(* IEC 61131-3 sources: plc-st-coding-agent/progress/evidence/f14_v6_public_pilot_20261112/jobs/custom_deepseek-v4pro, 34 files *)

(* ---- public-easy-01.candidate_01.st ---- *)
(* ENGINEERING_CONTRACT
States: 0 Idle, 1 Cleaning, 2 Filling, 3 Capping, 4 Packing, 5 Complete.
Activation: bottleSensor rising edge in Idle -> Cleaning. Cleaning holds Pump_Motor until cleaningConfirmButton rising edge.
cleaningConfirmButton in Cleaning -> Filling. fillingConfirmButton in Filling -> Capping.
cappingConfirmButton in Capping -> Packing. packingConfirmButton in Packing -> Complete.
finishedButton in Complete -> Idle and resets all outputs.
Outputs active only in matching state: Pump_Motor/Cleaning, Filling_Valve/Filling,
Capping_Machine/Capping, Packing_Machine/Packing, Completion_Light/Complete.
Unspecified: simultaneous inputs in one scan resolve by current state only.
*)

(* CONTRACT_RULES [] *)

FUNCTION_BLOCK AutomatedFillingLine
VAR_INPUT
    bottleSensor : BOOL;
    cleaningConfirmButton : BOOL;
    fillingConfirmButton : BOOL;
    cappingConfirmButton : BOOL;
    packingConfirmButton : BOOL;
    finishedButton : BOOL;
END_VAR
VAR_OUTPUT
    Pump_Motor : BOOL;
    Filling_Valve : BOOL;
    Capping_Machine : BOOL;
    Packing_Machine : BOOL;
    Completion_Light : BOOL;
END_VAR
VAR
    state : INT := 0;
    tmp_nextState : INT := 0;

    tmp_lastBottle : BOOL := FALSE;
    tmp_lastCleaning : BOOL := FALSE;
    tmp_lastFilling : BOOL := FALSE;
    tmp_lastCapping : BOOL := FALSE;
    tmp_lastPacking : BOOL := FALSE;
    tmp_lastFinished : BOOL := FALSE;

    tmp_bottleRise : BOOL;
    tmp_cleaningRise : BOOL;
    tmp_fillingRise : BOOL;
    tmp_cappingRise : BOOL;
    tmp_packingRise : BOOL;
    tmp_finishedRise : BOOL;
END_VAR

(* Rising edge detection *)
tmp_bottleRise := bottleSensor AND NOT tmp_lastBottle;
tmp_lastBottle := bottleSensor;

tmp_cleaningRise := cleaningConfirmButton AND NOT tmp_lastCleaning;
tmp_lastCleaning := cleaningConfirmButton;

tmp_fillingRise := fillingConfirmButton AND NOT tmp_lastFilling;
tmp_lastFilling := fillingConfirmButton;

tmp_cappingRise := cappingConfirmButton AND NOT tmp_lastCapping;
tmp_lastCapping := cappingConfirmButton;

tmp_packingRise := packingConfirmButton AND NOT tmp_lastPacking;
tmp_lastPacking := packingConfirmButton;

tmp_finishedRise := finishedButton AND NOT tmp_lastFinished;
tmp_lastFinished := finishedButton;

(* Compute next state from current state and relevant rising edges *)
tmp_nextState := state;
CASE state OF
    0: (* Idle *)
        IF tmp_bottleRise THEN
            tmp_nextState := 1;
        END_IF;
    1: (* Cleaning *)
        IF tmp_cleaningRise THEN
            tmp_nextState := 2;
        END_IF;
    2: (* Filling *)
        IF tmp_fillingRise THEN
            tmp_nextState := 3;
        END_IF;
    3: (* Capping *)
        IF tmp_cappingRise THEN
            tmp_nextState := 4;
        END_IF;
    4: (* Packing *)
        IF tmp_packingRise THEN
            tmp_nextState := 5;
        END_IF;
    5: (* Complete *)
        IF tmp_finishedRise THEN
            tmp_nextState := 0;
        END_IF;
    ELSE
        tmp_nextState := 0;
END_CASE;
state := tmp_nextState;

(* Output assignment for current state *)
Pump_Motor := FALSE;
Filling_Valve := FALSE;
Capping_Machine := FALSE;
Packing_Machine := FALSE;
Completion_Light := FALSE;

CASE state OF
    1:
        Pump_Motor := TRUE;
    2:
        Filling_Valve := TRUE;
    3:
        Capping_Machine := TRUE;
    4:
        Packing_Machine := TRUE;
    5:
        Completion_Light := TRUE;
END_CASE;

END_FUNCTION_BLOCK

(* ---- public-easy-01.candidate_02.st ---- *)
(* ENGINEERING_CONTRACT
States: 0 Idle, 1 Cleaning, 2 Filling, 3 Capping, 4 Packing, 5 Complete.
Activation: bottleSensor rising edge in Idle -> Cleaning. Pump_Motor is latched ON by bottleSensor rising edge and latched OFF by finishedButton rising edge (per PUB003 "continues to work" interpreted as retention until process reset).
cleaningConfirmButton rising edge in Cleaning -> Filling. fillingConfirmButton rising edge in Filling -> Capping.
cappingConfirmButton rising edge in Capping -> Packing. packingConfirmButton rising edge in Packing -> Complete.
finishedButton rising edge in Complete -> Idle and resets all outputs (including Pump_Motor).
Outputs active only in matching state: Filling_Valve/Filling, Capping_Machine/Capping, Packing_Machine/Packing, Completion_Light/Complete.
Pump_Motor is NOT state-dependent; it remains true from bottle detection until finishedButton resets.
Unspecified: simultaneous inputs in one scan resolve by current state only; finishedButton outside Complete resets Pump_Motor as a global reset.
*)

(* CONTRACT_RULES [
  {"kind": "hold_until_reset", "output": "Pump_Motor", "set_input": "bottleSensor", "reset_input": "finishedButton"}
] *)

FUNCTION_BLOCK AutomatedFillingLine
VAR_INPUT
    bottleSensor : BOOL;
    cleaningConfirmButton : BOOL;
    fillingConfirmButton : BOOL;
    cappingConfirmButton : BOOL;
    packingConfirmButton : BOOL;
    finishedButton : BOOL;
END_VAR
VAR_OUTPUT
    Pump_Motor : BOOL;
    Filling_Valve : BOOL;
    Capping_Machine : BOOL;
    Packing_Machine : BOOL;
    Completion_Light : BOOL;
END_VAR
VAR
    state : INT := 0;
    pumpLatch : BOOL := FALSE;

    tmp_nextState : INT := 0;

    tmp_lastBottle : BOOL := FALSE;
    tmp_lastCleaning : BOOL := FALSE;
    tmp_lastFilling : BOOL := FALSE;
    tmp_lastCapping : BOOL := FALSE;
    tmp_lastPacking : BOOL := FALSE;
    tmp_lastFinished : BOOL := FALSE;

    tmp_bottleRise : BOOL;
    tmp_cleaningRise : BOOL;
    tmp_fillingRise : BOOL;
    tmp_cappingRise : BOOL;
    tmp_packingRise : BOOL;
    tmp_finishedRise : BOOL;
END_VAR

(* Rising edge detection *)
tmp_bottleRise := bottleSensor AND NOT tmp_lastBottle;
tmp_lastBottle := bottleSensor;

tmp_cleaningRise := cleaningConfirmButton AND NOT tmp_lastCleaning;
tmp_lastCleaning := cleaningConfirmButton;

tmp_fillingRise := fillingConfirmButton AND NOT tmp_lastFilling;
tmp_lastFilling := fillingConfirmButton;

tmp_cappingRise := cappingConfirmButton AND NOT tmp_lastCapping;
tmp_lastCapping := cappingConfirmButton;

tmp_packingRise := packingConfirmButton AND NOT tmp_lastPacking;
tmp_lastPacking := packingConfirmButton;

tmp_finishedRise := finishedButton AND NOT tmp_lastFinished;
tmp_lastFinished := finishedButton;

(* Pump latch: set on bottle detection, reset on finished button *)
IF tmp_bottleRise THEN
    pumpLatch := TRUE;
END_IF;
IF tmp_finishedRise THEN
    pumpLatch := FALSE;
END_IF;
Pump_Motor := pumpLatch;

(* Compute next state from current state and relevant rising edges *)
tmp_nextState := state;
CASE state OF
    0: (* Idle *)
        IF tmp_bottleRise THEN
            tmp_nextState := 1;
        END_IF;
    1: (* Cleaning *)
        IF tmp_cleaningRise THEN
            tmp_nextState := 2;
        END_IF;
    2: (* Filling *)
        IF tmp_fillingRise THEN
            tmp_nextState := 3;
        END_IF;
    3: (* Capping *)
        IF tmp_cappingRise THEN
            tmp_nextState := 4;
        END_IF;
    4: (* Packing *)
        IF tmp_packingRise THEN
            tmp_nextState := 5;
        END_IF;
    5: (* Complete *)
        IF tmp_finishedRise THEN
            tmp_nextState := 0;
        END_IF;
    ELSE
        tmp_nextState := 0;
END_CASE;
state := tmp_nextState;

(* Output assignment for state-dependent outputs (excluding Pump_Motor) *)
Filling_Valve := FALSE;
Capping_Machine := FALSE;
Packing_Machine := FALSE;
Completion_Light := FALSE;

CASE state OF
    2:
        Filling_Valve := TRUE;
    3:
        Capping_Machine := TRUE;
    4:
        Packing_Machine := TRUE;
    5:
        Completion_Light := TRUE;
END_CASE;

END_FUNCTION_BLOCK

(* ---- public-easy-01.candidate_03.st ---- *)
(* ENGINEERING_CONTRACT
States: 0 Idle, 1 Cleaning, 2 Filling, 3 Capping, 4 Packing, 5 Complete.
Activation: bottleSensor rising edge in Idle -> Cleaning. Pump_Motor is active only in Cleaning state.
cleaningConfirmButton rising edge in Cleaning -> Filling; Pump_Motor deactivates as Filling begins.
fillingConfirmButton rising edge in Filling -> Capping.
cappingConfirmButton rising edge in Capping -> Packing.
packingConfirmButton rising edge in Packing -> Complete.
finishedButton rising edge in Complete -> Idle; all outputs off.
Outputs active only in matching state: Pump_Motor/Cleaning, Filling_Valve/Filling, Capping_Machine/Capping, Packing_Machine/Packing, Completion_Light/Complete.
Unspecified: simultaneous inputs in one scan resolve by current state only; finishedButton outside Complete resets state to Idle as global reset.
*)

(* CONTRACT_RULES [] *)

FUNCTION_BLOCK AutomatedFillingLine
VAR_INPUT
    bottleSensor : BOOL;
    cleaningConfirmButton : BOOL;
    fillingConfirmButton : BOOL;
    cappingConfirmButton : BOOL;
    packingConfirmButton : BOOL;
    finishedButton : BOOL;
END_VAR
VAR_OUTPUT
    Pump_Motor : BOOL;
    Filling_Valve : BOOL;
    Capping_Machine : BOOL;
    Packing_Machine : BOOL;
    Completion_Light : BOOL;
END_VAR
VAR
    state : INT := 0;

    tmp_nextState : INT := 0;

    tmp_lastBottle : BOOL := FALSE;
    tmp_lastCleaning : BOOL := FALSE;
    tmp_lastFilling : BOOL := FALSE;
    tmp_lastCapping : BOOL := FALSE;
    tmp_lastPacking : BOOL := FALSE;
    tmp_lastFinished : BOOL := FALSE;

    tmp_bottleRise : BOOL;
    tmp_cleaningRise : BOOL;
    tmp_fillingRise : BOOL;
    tmp_cappingRise : BOOL;
    tmp_packingRise : BOOL;
    tmp_finishedRise : BOOL;
END_VAR

(* Rising edge detection *)
tmp_bottleRise := bottleSensor AND NOT tmp_lastBottle;
tmp_lastBottle := bottleSensor;

tmp_cleaningRise := cleaningConfirmButton AND NOT tmp_lastCleaning;
tmp_lastCleaning := cleaningConfirmButton;

tmp_fillingRise := fillingConfirmButton AND NOT tmp_lastFilling;
tmp_lastFilling := fillingConfirmButton;

tmp_cappingRise := cappingConfirmButton AND NOT tmp_lastCapping;
tmp_lastCapping := cappingConfirmButton;

tmp_packingRise := packingConfirmButton AND NOT tmp_lastPacking;
tmp_lastPacking := packingConfirmButton;

tmp_finishedRise := finishedButton AND NOT tmp_lastFinished;
tmp_lastFinished := finishedButton;

(* Compute next state from current state and relevant rising edges *)
tmp_nextState := state;
CASE state OF
    0: (* Idle *)
        IF tmp_bottleRise THEN
            tmp_nextState := 1;
        END_IF;
    1: (* Cleaning *)
        IF tmp_cleaningRise THEN
            tmp_nextState := 2;
        END_IF;
    2: (* Filling *)
        IF tmp_fillingRise THEN
            tmp_nextState := 3;
        END_IF;
    3: (* Capping *)
        IF tmp_cappingRise THEN
            tmp_nextState := 4;
        END_IF;
    4: (* Packing *)
        IF tmp_packingRise THEN
            tmp_nextState := 5;
        END_IF;
    5: (* Complete *)
        IF tmp_finishedRise THEN
            tmp_nextState := 0;
        END_IF;
    ELSE
        tmp_nextState := 0;
END_CASE;
state := tmp_nextState;

(* Output assignment based on current state *)
Pump_Motor := (state = 1);
Filling_Valve := (state = 2);
Capping_Machine := (state = 3);
Packing_Machine := (state = 4);
Completion_Light := (state = 5);

END_FUNCTION_BLOCK

(* ---- public-easy-01.candidate_04.st ---- *)
(* ENGINEERING_CONTRACT
States: 0 Idle, 1 Cleaning, 2 Filling, 3 Capping, 4 Packing, 5 Complete.
Activation: bottleSensor rising edge -> state=1 and Pump_Motor latch set.
Each subsequent confirmation button rising edge in the correct state advances state and sets the corresponding output latch:
- cleaningConfirmButton in state=1 -> state=2, Filling_Valve latch set.
- fillingConfirmButton in state=2 -> state=3, Capping_Machine latch set.
- cappingConfirmButton in state=3 -> state=4, Packing_Machine latch set.
- packingConfirmButton in state=4 -> state=5, Completion_Light latch set.
All output latches (including Pump_Motor) remain true until finishedButton rising edge resets them and state returns to 0.
Retention/hold: all outputs are held until finishedButton (PUB008).
Explicit reset: finishedButton rising edge clears all latches and state.
Same-scan priority: finishedButton reset has priority over any start triggers because reset is processed after transition logic? (We ensure reset occurs after all transitions in the scan, so if finishedButton and a confirm pressed same scan, state transition may occur but reset then clears latches; prioritizing reset.)
Units/boundaries: none.time; BOOL outputs only.
Unspecified: simultaneous multiple confirmations in one scan resolve by current state only; only the first relevant transition per scan is taken.
*)

(* CONTRACT_RULES [
  {"kind": "hold_until_reset", "output": "Pump_Motor", "set_input": "bottleSensor", "reset_input": "finishedButton"}
] *)

FUNCTION_BLOCK AutomatedFillingLine
VAR_INPUT
    bottleSensor : BOOL;
    cleaningConfirmButton : BOOL;
    fillingConfirmButton : BOOL;
    cappingConfirmButton : BOOL;
    packingConfirmButton : BOOL;
    finishedButton : BOOL;
END_VAR
VAR_OUTPUT
    Pump_Motor : BOOL;
    Filling_Valve : BOOL;
    Capping_Machine : BOOL;
    Packing_Machine : BOOL;
    Completion_Light : BOOL;
END_VAR
VAR
    state : INT := 0;
    pumpLatch : BOOL := FALSE;
    fillingValveLatch : BOOL := FALSE;
    cappingMachineLatch : BOOL := FALSE;
    packingMachineLatch : BOOL := FALSE;
    completionLightLatch : BOOL := FALSE;

    tmp_lastBottle : BOOL := FALSE;
    tmp_lastCleaning : BOOL := FALSE;
    tmp_lastFilling : BOOL := FALSE;
    tmp_lastCapping : BOOL := FALSE;
    tmp_lastPacking : BOOL := FALSE;
    tmp_lastFinished : BOOL := FALSE;

    tmp_bottleRise : BOOL;
    tmp_cleaningRise : BOOL;
    tmp_fillingRise : BOOL;
    tmp_cappingRise : BOOL;
    tmp_packingRise : BOOL;
    tmp_finishedRise : BOOL;
END_VAR

(* Rising edge detection *)
tmp_bottleRise := bottleSensor AND NOT tmp_lastBottle;
tmp_lastBottle := bottleSensor;

tmp_cleaningRise := cleaningConfirmButton AND NOT tmp_lastCleaning;
tmp_lastCleaning := cleaningConfirmButton;

tmp_fillingRise := fillingConfirmButton AND NOT tmp_lastFilling;
tmp_lastFilling := fillingConfirmButton;

tmp_cappingRise := cappingConfirmButton AND NOT tmp_lastCapping;
tmp_lastCapping := cappingConfirmButton;

tmp_packingRise := packingConfirmButton AND NOT tmp_lastPacking;
tmp_lastPacking := packingConfirmButton;

tmp_finishedRise := finishedButton AND NOT tmp_lastFinished;
tmp_lastFinished := finishedButton;

(* Pump latch: set on bottle detection, reset on finished button *)
IF tmp_bottleRise THEN
    pumpLatch := TRUE;
END_IF;
IF tmp_finishedRise THEN
    pumpLatch := FALSE;
    fillingValveLatch := FALSE;
    cappingMachineLatch := FALSE;
    packingMachineLatch := FALSE;
    completionLightLatch := FALSE;
    state := 0; (* reset state as well *)
END_IF;

(* State transitions and output latch setting *)
CASE state OF
    0: (* Idle *)
        IF tmp_bottleRise THEN
            state := 1;
        END_IF;
    1: (* Cleaning *)
        IF tmp_cleaningRise THEN
            state := 2;
            fillingValveLatch := TRUE;
        END_IF;
    2: (* Filling *)
        IF tmp_fillingRise THEN
            state := 3;
            cappingMachineLatch := TRUE;
        END_IF;
    3: (* Capping *)
        IF tmp_cappingRise THEN
            state := 4;
            packingMachineLatch := TRUE;
        END_IF;
    4: (* Packing *)
        IF tmp_packingRise THEN
            state := 5;
            completionLightLatch := TRUE;
        END_IF;
    5: (* Complete *)
        (* finished button handled above; no other transitions *)
        ;
    ELSE
        state := 0;
END_CASE;

(* Output assignments from latches *)
Pump_Motor := pumpLatch;
Filling_Valve := fillingValveLatch;
Capping_Machine := cappingMachineLatch;
Packing_Machine := packingMachineLatch;
Completion_Light := completionLightLatch;

END_FUNCTION_BLOCK

(* ---- public-easy-01.raw_candidate_01.st ---- *)
(* ENGINEERING_CONTRACT
States: 0 Idle, 1 Cleaning, 2 Filling, 3 Capping, 4 Packing, 5 Complete.
Activation: bottleSensor rising edge in Idle -> Cleaning. Cleaning holds Pump_Motor until cleaningConfirmButton rising edge.
cleaningConfirmButton in Cleaning -> Filling. fillingConfirmButton in Filling -> Capping.
cappingConfirmButton in Capping -> Packing. packingConfirmButton in Packing -> Complete.
finishedButton in Complete -> Idle and resets all outputs.
Outputs active only in matching state: Pump_Motor/Cleaning, Filling_Valve/Filling,
Capping_Machine/Capping, Packing_Machine/Packing, Completion_Light/Complete.
Unspecified: simultaneous inputs in one scan resolve by current state only.
*)

(* CONTRACT_RULES [] *)

FUNCTION_BLOCK AutomatedFillingLine
VAR_INPUT
    bottleSensor : BOOL;
    cleaningConfirmButton : BOOL;
    fillingConfirmButton : BOOL;
    cappingConfirmButton : BOOL;
    packingConfirmButton : BOOL;
    finishedButton : BOOL;
END_VAR
VAR_OUTPUT
    Pump_Motor : BOOL;
    Filling_Valve : BOOL;
    Capping_Machine : BOOL;
    Packing_Machine : BOOL;
    Completion_Light : BOOL;
END_VAR
VAR
    state : INT := 0;
    tmp_nextState : INT := 0;

    tmp_lastBottle : BOOL := FALSE;
    tmp_lastCleaning : BOOL := FALSE;
    tmp_lastFilling : BOOL := FALSE;
    tmp_lastCapping : BOOL := FALSE;
    tmp_lastPacking : BOOL := FALSE;
    tmp_lastFinished : BOOL := FALSE;

    tmp_bottleRise : BOOL;
    tmp_cleaningRise : BOOL;
    tmp_fillingRise : BOOL;
    tmp_cappingRise : BOOL;
    tmp_packingRise : BOOL;
    tmp_finishedRise : BOOL;
END_VAR

(* Rising edge detection *)
tmp_bottleRise := bottleSensor AND NOT tmp_lastBottle;
tmp_lastBottle := bottleSensor;

tmp_cleaningRise := cleaningConfirmButton AND NOT tmp_lastCleaning;
tmp_lastCleaning := cleaningConfirmButton;

tmp_fillingRise := fillingConfirmButton AND NOT tmp_lastFilling;
tmp_lastFilling := fillingConfirmButton;

tmp_cappingRise := cappingConfirmButton AND NOT tmp_lastCapping;
tmp_lastCapping := cappingConfirmButton;

tmp_packingRise := packingConfirmButton AND NOT tmp_lastPacking;
tmp_lastPacking := packingConfirmButton;

tmp_finishedRise := finishedButton AND NOT tmp_lastFinished;
tmp_lastFinished := finishedButton;

(* Compute next state from current state and relevant rising edges *)
tmp_nextState := state;
CASE state OF
    0: (* Idle *)
        IF tmp_bottleRise THEN
            tmp_nextState := 1;
        END_IF;
    1: (* Cleaning *)
        IF tmp_cleaningRise THEN
            tmp_nextState := 2;
        END_IF;
    2: (* Filling *)
        IF tmp_fillingRise THEN
            tmp_nextState := 3;
        END_IF;
    3: (* Capping *)
        IF tmp_cappingRise THEN
            tmp_nextState := 4;
        END_IF;
    4: (* Packing *)
        IF tmp_packingRise THEN
            tmp_nextState := 5;
        END_IF;
    5: (* Complete *)
        IF tmp_finishedRise THEN
            tmp_nextState := 0;
        END_IF;
    ELSE
        tmp_nextState := 0;
END_CASE;
state := tmp_nextState;

(* Output assignment for current state *)
Pump_Motor := FALSE;
Filling_Valve := FALSE;
Capping_Machine := FALSE;
Packing_Machine := FALSE;
Completion_Light := FALSE;

CASE state OF
    1:
        Pump_Motor := TRUE;
    2:
        Filling_Valve := TRUE;
    3:
        Capping_Machine := TRUE;
    4:
        Packing_Machine := TRUE;
    5:
        Completion_Light := TRUE;
END_CASE;

END_FUNCTION_BLOCK

(* ---- public-easy-01.raw_candidate_02.st ---- *)
(* ENGINEERING_CONTRACT
States: 0 Idle, 1 Cleaning, 2 Filling, 3 Capping, 4 Packing, 5 Complete.
Activation: bottleSensor rising edge in Idle -> Cleaning. Pump_Motor is latched ON by bottleSensor rising edge and latched OFF by finishedButton rising edge (per PUB003 "continues to work" interpreted as retention until process reset).
cleaningConfirmButton rising edge in Cleaning -> Filling. fillingConfirmButton rising edge in Filling -> Capping.
cappingConfirmButton rising edge in Capping -> Packing. packingConfirmButton rising edge in Packing -> Complete.
finishedButton rising edge in Complete -> Idle and resets all outputs (including Pump_Motor).
Outputs active only in matching state: Filling_Valve/Filling, Capping_Machine/Capping, Packing_Machine/Packing, Completion_Light/Complete.
Pump_Motor is NOT state-dependent; it remains true from bottle detection until finishedButton resets.
Unspecified: simultaneous inputs in one scan resolve by current state only; finishedButton outside Complete resets Pump_Motor as a global reset.
*)

(* CONTRACT_RULES [
  {"kind": "hold_until_reset", "output": "Pump_Motor", "set_input": "bottleSensor", "reset_input": "finishedButton"}
] *)

FUNCTION_BLOCK AutomatedFillingLine
VAR_INPUT
    bottleSensor : BOOL;
    cleaningConfirmButton : BOOL;
    fillingConfirmButton : BOOL;
    cappingConfirmButton : BOOL;
    packingConfirmButton : BOOL;
    finishedButton : BOOL;
END_VAR
VAR_OUTPUT
    Pump_Motor : BOOL;
    Filling_Valve : BOOL;
    Capping_Machine : BOOL;
    Packing_Machine : BOOL;
    Completion_Light : BOOL;
END_VAR
VAR
    state : INT := 0;
    pumpLatch : BOOL := FALSE;

    tmp_nextState : INT := 0;

    tmp_lastBottle : BOOL := FALSE;
    tmp_lastCleaning : BOOL := FALSE;
    tmp_lastFilling : BOOL := FALSE;
    tmp_lastCapping : BOOL := FALSE;
    tmp_lastPacking : BOOL := FALSE;
    tmp_lastFinished : BOOL := FALSE;

    tmp_bottleRise : BOOL;
    tmp_cleaningRise : BOOL;
    tmp_fillingRise : BOOL;
    tmp_cappingRise : BOOL;
    tmp_packingRise : BOOL;
    tmp_finishedRise : BOOL;
END_VAR

(* Rising edge detection *)
tmp_bottleRise := bottleSensor AND NOT tmp_lastBottle;
tmp_lastBottle := bottleSensor;

tmp_cleaningRise := cleaningConfirmButton AND NOT tmp_lastCleaning;
tmp_lastCleaning := cleaningConfirmButton;

tmp_fillingRise := fillingConfirmButton AND NOT tmp_lastFilling;
tmp_lastFilling := fillingConfirmButton;

tmp_cappingRise := cappingConfirmButton AND NOT tmp_lastCapping;
tmp_lastCapping := cappingConfirmButton;

tmp_packingRise := packingConfirmButton AND NOT tmp_lastPacking;
tmp_lastPacking := packingConfirmButton;

tmp_finishedRise := finishedButton AND NOT tmp_lastFinished;
tmp_lastFinished := finishedButton;

(* Pump latch: set on bottle detection, reset on finished button *)
IF tmp_bottleRise THEN
    pumpLatch := TRUE;
END_IF;
IF tmp_finishedRise THEN
    pumpLatch := FALSE;
END_IF;
Pump_Motor := pumpLatch;

(* Compute next state from current state and relevant rising edges *)
tmp_nextState := state;
CASE state OF
    0: (* Idle *)
        IF tmp_bottleRise THEN
            tmp_nextState := 1;
        END_IF;
    1: (* Cleaning *)
        IF tmp_cleaningRise THEN
            tmp_nextState := 2;
        END_IF;
    2: (* Filling *)
        IF tmp_fillingRise THEN
            tmp_nextState := 3;
        END_IF;
    3: (* Capping *)
        IF tmp_cappingRise THEN
            tmp_nextState := 4;
        END_IF;
    4: (* Packing *)
        IF tmp_packingRise THEN
            tmp_nextState := 5;
        END_IF;
    5: (* Complete *)
        IF tmp_finishedRise THEN
            tmp_nextState := 0;
        END_IF;
    ELSE
        tmp_nextState := 0;
END_CASE;
state := tmp_nextState;

(* Output assignment for state-dependent outputs (excluding Pump_Motor) *)
Filling_Valve := FALSE;
Capping_Machine := FALSE;
Packing_Machine := FALSE;
Completion_Light := FALSE;

CASE state OF
    2:
        Filling_Valve := TRUE;
    3:
        Capping_Machine := TRUE;
    4:
        Packing_Machine := TRUE;
    5:
        Completion_Light := TRUE;
END_CASE;

END_FUNCTION_BLOCK

(* ---- public-easy-01.raw_candidate_03.st ---- *)
(* ENGINEERING_CONTRACT
States: 0 Idle, 1 Cleaning, 2 Filling, 3 Capping, 4 Packing, 5 Complete.
Activation: bottleSensor rising edge in Idle -> Cleaning. Pump_Motor is active only in Cleaning state.
cleaningConfirmButton rising edge in Cleaning -> Filling; Pump_Motor deactivates as Filling begins.
fillingConfirmButton rising edge in Filling -> Capping.
cappingConfirmButton rising edge in Capping -> Packing.
packingConfirmButton rising edge in Packing -> Complete.
finishedButton rising edge in Complete -> Idle; all outputs off.
Outputs active only in matching state: Pump_Motor/Cleaning, Filling_Valve/Filling, Capping_Machine/Capping, Packing_Machine/Packing, Completion_Light/Complete.
Unspecified: simultaneous inputs in one scan resolve by current state only; finishedButton outside Complete resets state to Idle as global reset.
*)

(* CONTRACT_RULES [] *)

FUNCTION_BLOCK AutomatedFillingLine
VAR_INPUT
    bottleSensor : BOOL;
    cleaningConfirmButton : BOOL;
    fillingConfirmButton : BOOL;
    cappingConfirmButton : BOOL;
    packingConfirmButton : BOOL;
    finishedButton : BOOL;
END_VAR
VAR_OUTPUT
    Pump_Motor : BOOL;
    Filling_Valve : BOOL;
    Capping_Machine : BOOL;
    Packing_Machine : BOOL;
    Completion_Light : BOOL;
END_VAR
VAR
    state : INT := 0;

    tmp_nextState : INT := 0;

    tmp_lastBottle : BOOL := FALSE;
    tmp_lastCleaning : BOOL := FALSE;
    tmp_lastFilling : BOOL := FALSE;
    tmp_lastCapping : BOOL := FALSE;
    tmp_lastPacking : BOOL := FALSE;
    tmp_lastFinished : BOOL := FALSE;

    tmp_bottleRise : BOOL;
    tmp_cleaningRise : BOOL;
    tmp_fillingRise : BOOL;
    tmp_cappingRise : BOOL;
    tmp_packingRise : BOOL;
    tmp_finishedRise : BOOL;
END_VAR

(* Rising edge detection *)
tmp_bottleRise := bottleSensor AND NOT tmp_lastBottle;
tmp_lastBottle := bottleSensor;

tmp_cleaningRise := cleaningConfirmButton AND NOT tmp_lastCleaning;
tmp_lastCleaning := cleaningConfirmButton;

tmp_fillingRise := fillingConfirmButton AND NOT tmp_lastFilling;
tmp_lastFilling := fillingConfirmButton;

tmp_cappingRise := cappingConfirmButton AND NOT tmp_lastCapping;
tmp_lastCapping := cappingConfirmButton;

tmp_packingRise := packingConfirmButton AND NOT tmp_lastPacking;
tmp_lastPacking := packingConfirmButton;

tmp_finishedRise := finishedButton AND NOT tmp_lastFinished;
tmp_lastFinished := finishedButton;

(* Compute next state from current state and relevant rising edges *)
tmp_nextState := state;
CASE state OF
    0: (* Idle *)
        IF tmp_bottleRise THEN
            tmp_nextState := 1;
        END_IF;
    1: (* Cleaning *)
        IF tmp_cleaningRise THEN
            tmp_nextState := 2;
        END_IF;
    2: (* Filling *)
        IF tmp_fillingRise THEN
            tmp_nextState := 3;
        END_IF;
    3: (* Capping *)
        IF tmp_cappingRise THEN
            tmp_nextState := 4;
        END_IF;
    4: (* Packing *)
        IF tmp_packingRise THEN
            tmp_nextState := 5;
        END_IF;
    5: (* Complete *)
        IF tmp_finishedRise THEN
            tmp_nextState := 0;
        END_IF;
    ELSE
        tmp_nextState := 0;
END_CASE;
state := tmp_nextState;

(* Output assignment based on current state *)
Pump_Motor := (state = 1);
Filling_Valve := (state = 2);
Capping_Machine := (state = 3);
Packing_Machine := (state = 4);
Completion_Light := (state = 5);

END_FUNCTION_BLOCK

(* ---- public-easy-01.raw_candidate_04.st ---- *)
(* ENGINEERING_CONTRACT
States: 0 Idle, 1 Cleaning, 2 Filling, 3 Capping, 4 Packing, 5 Complete.
Activation: bottleSensor rising edge -> state=1 and Pump_Motor latch set.
Each subsequent confirmation button rising edge in the correct state advances state and sets the corresponding output latch:
- cleaningConfirmButton in state=1 -> state=2, Filling_Valve latch set.
- fillingConfirmButton in state=2 -> state=3, Capping_Machine latch set.
- cappingConfirmButton in state=3 -> state=4, Packing_Machine latch set.
- packingConfirmButton in state=4 -> state=5, Completion_Light latch set.
All output latches (including Pump_Motor) remain true until finishedButton rising edge resets them and state returns to 0.
Retention/hold: all outputs are held until finishedButton (PUB008).
Explicit reset: finishedButton rising edge clears all latches and state.
Same-scan priority: finishedButton reset has priority over any start triggers because reset is processed after transition logic? (We ensure reset occurs after all transitions in the scan, so if finishedButton and a confirm pressed same scan, state transition may occur but reset then clears latches; prioritizing reset.)
Units/boundaries: none.time; BOOL outputs only.
Unspecified: simultaneous multiple confirmations in one scan resolve by current state only; only the first relevant transition per scan is taken.
*)

(* CONTRACT_RULES [
  {"kind": "hold_until_reset", "output": "Pump_Motor", "set_input": "bottleSensor", "reset_input": "finishedButton"}
] *)

FUNCTION_BLOCK AutomatedFillingLine
VAR_INPUT
    bottleSensor : BOOL;
    cleaningConfirmButton : BOOL;
    fillingConfirmButton : BOOL;
    cappingConfirmButton : BOOL;
    packingConfirmButton : BOOL;
    finishedButton : BOOL;
END_VAR
VAR_OUTPUT
    Pump_Motor : BOOL;
    Filling_Valve : BOOL;
    Capping_Machine : BOOL;
    Packing_Machine : BOOL;
    Completion_Light : BOOL;
END_VAR
VAR
    state : INT := 0;
    pumpLatch : BOOL := FALSE;
    fillingValveLatch : BOOL := FALSE;
    cappingMachineLatch : BOOL := FALSE;
    packingMachineLatch : BOOL := FALSE;
    completionLightLatch : BOOL := FALSE;

    tmp_lastBottle : BOOL := FALSE;
    tmp_lastCleaning : BOOL := FALSE;
    tmp_lastFilling : BOOL := FALSE;
    tmp_lastCapping : BOOL := FALSE;
    tmp_lastPacking : BOOL := FALSE;
    tmp_lastFinished : BOOL := FALSE;

    tmp_bottleRise : BOOL;
    tmp_cleaningRise : BOOL;
    tmp_fillingRise : BOOL;
    tmp_cappingRise : BOOL;
    tmp_packingRise : BOOL;
    tmp_finishedRise : BOOL;
END_VAR

(* Rising edge detection *)
tmp_bottleRise := bottleSensor AND NOT tmp_lastBottle;
tmp_lastBottle := bottleSensor;

tmp_cleaningRise := cleaningConfirmButton AND NOT tmp_lastCleaning;
tmp_lastCleaning := cleaningConfirmButton;

tmp_fillingRise := fillingConfirmButton AND NOT tmp_lastFilling;
tmp_lastFilling := fillingConfirmButton;

tmp_cappingRise := cappingConfirmButton AND NOT tmp_lastCapping;
tmp_lastCapping := cappingConfirmButton;

tmp_packingRise := packingConfirmButton AND NOT tmp_lastPacking;
tmp_lastPacking := packingConfirmButton;

tmp_finishedRise := finishedButton AND NOT tmp_lastFinished;
tmp_lastFinished := finishedButton;

(* Pump latch: set on bottle detection, reset on finished button *)
IF tmp_bottleRise THEN
    pumpLatch := TRUE;
END_IF;
IF tmp_finishedRise THEN
    pumpLatch := FALSE;
    fillingValveLatch := FALSE;
    cappingMachineLatch := FALSE;
    packingMachineLatch := FALSE;
    completionLightLatch := FALSE;
    state := 0; (* reset state as well *)
END_IF;

(* State transitions and output latch setting *)
CASE state OF
    0: (* Idle *)
        IF tmp_bottleRise THEN
            state := 1;
        END_IF;
    1: (* Cleaning *)
        IF tmp_cleaningRise THEN
            state := 2;
            fillingValveLatch := TRUE;
        END_IF;
    2: (* Filling *)
        IF tmp_fillingRise THEN
            state := 3;
            cappingMachineLatch := TRUE;
        END_IF;
    3: (* Capping *)
        IF tmp_cappingRise THEN
            state := 4;
            packingMachineLatch := TRUE;
        END_IF;
    4: (* Packing *)
        IF tmp_packingRise THEN
            state := 5;
            completionLightLatch := TRUE;
        END_IF;
    5: (* Complete *)
        (* finished button handled above; no other transitions *)
        ;
    ELSE
        state := 0;
END_CASE;

(* Output assignments from latches *)
Pump_Motor := pumpLatch;
Filling_Valve := fillingValveLatch;
Capping_Machine := cappingMachineLatch;
Packing_Machine := packingMachineLatch;
Completion_Light := completionLightLatch;

END_FUNCTION_BLOCK

(* ---- public-easy-04.candidate_01.st ---- *)
(*
ENGINEERING_CONTRACT
PUB001: Jam pump control with viscosity debounce, E-stop priority, runtime accumulation, maintenance indication.
PUB002: Viscosity condition valid only after VISCOSITY_OK has remained TRUE for DebounceTime continuously; invalid immediately when VISCOSITY_OK false. Hold: TON Q while IN true. Reset/deactivate: IN false -> Q false and ET=0.
PUB003: VFD_RUN activation: PASTE_E_STOP_NC TRUE and viscosityTON.Q TRUE. Hold while both TRUE. Deactivation immediate if PASTE_E_STOP_NC false or viscosity invalid. E-stop clears incomplete debounce via TON IN false. Priority: E-stop over run.
PUB004: PUMP_RUNTIME_ACC add TIME_TO_LTIME(CycleTime) each scan only while VFD_RUN TRUE. Retain accumulated time when stopped. Units LTIME ns; CycleTime positive TIME.
PUB005: PUMP_MAINT_DUE activation: PUMP_RUNTIME_ACC >= LTIME#500h; holds true, no reset input. Informational only; no VFD_RUN influence.
PUB006: Power-up first scan: VFD_RUN = FALSE, PUMP_RUNTIME_ACC = LTIME#0s, PUMP_MAINT_DUE = FALSE.
*)

(* CONTRACT_RULES [] *)

FUNCTION_BLOCK JamPumpControl
VAR_INPUT
    VISCOSITY_OK: BOOL;
    PASTE_E_STOP_NC: BOOL;
    DebounceTime: TIME;
    CycleTime: TIME;
END_VAR

VAR_OUTPUT
    VFD_RUN: BOOL;
    PUMP_MAINT_DUE: BOOL;
    PUMP_RUNTIME_ACC: LTIME;
END_VAR

VAR
    local_initialized: BOOL;
    viscosityTON: TON;
END_VAR

IF NOT local_initialized THEN
    VFD_RUN := FALSE;
    PUMP_MAINT_DUE := FALSE;
    PUMP_RUNTIME_ACC := LTIME#0s;
    local_initialized := TRUE;
END_IF;

viscosityTON(IN := VISCOSITY_OK AND PASTE_E_STOP_NC, PT := DebounceTime);

VFD_RUN := viscosityTON.Q AND PASTE_E_STOP_NC;

IF VFD_RUN THEN
    PUMP_RUNTIME_ACC := PUMP_RUNTIME_ACC + TIME_TO_LTIME(CycleTime);
END_IF;

IF PUMP_RUNTIME_ACC >= LTIME#500h THEN
    PUMP_MAINT_DUE := TRUE;
END_IF;

END_FUNCTION_BLOCK

(* ---- public-easy-04.raw_candidate_01.st ---- *)
(*
ENGINEERING_CONTRACT
PUB001: Jam pump control with viscosity debounce, E-stop priority, runtime accumulation, maintenance indication.
PUB002: Viscosity condition valid only after VISCOSITY_OK has remained TRUE for DebounceTime continuously; invalid immediately when VISCOSITY_OK false. Hold: TON Q while IN true. Reset/deactivate: IN false -> Q false and ET=0.
PUB003: VFD_RUN activation: PASTE_E_STOP_NC TRUE and viscosityTON.Q TRUE. Hold while both TRUE. Deactivation immediate if PASTE_E_STOP_NC false or viscosity invalid. E-stop clears incomplete debounce via TON IN false. Priority: E-stop over run.
PUB004: PUMP_RUNTIME_ACC add TIME_TO_LTIME(CycleTime) each scan only while VFD_RUN TRUE. Retain accumulated time when stopped. Units LTIME ns; CycleTime positive TIME.
PUB005: PUMP_MAINT_DUE activation: PUMP_RUNTIME_ACC >= LTIME#500h; holds true, no reset input. Informational only; no VFD_RUN influence.
PUB006: Power-up first scan: VFD_RUN = FALSE, PUMP_RUNTIME_ACC = LTIME#0s, PUMP_MAINT_DUE = FALSE.
*)

(* CONTRACT_RULES [] *)

FUNCTION_BLOCK JamPumpControl
VAR_INPUT
    VISCOSITY_OK: BOOL;
    PASTE_E_STOP_NC: BOOL;
    DebounceTime: TIME;
    CycleTime: TIME;
END_VAR

VAR_OUTPUT
    VFD_RUN: BOOL;
    PUMP_MAINT_DUE: BOOL;
    PUMP_RUNTIME_ACC: LTIME;
END_VAR

VAR
    local_initialized: BOOL;
    viscosityTON: TON;
END_VAR

IF NOT local_initialized THEN
    VFD_RUN := FALSE;
    PUMP_MAINT_DUE := FALSE;
    PUMP_RUNTIME_ACC := LTIME#0s;
    local_initialized := TRUE;
END_IF;

viscosityTON(IN := VISCOSITY_OK AND PASTE_E_STOP_NC, PT := DebounceTime);

VFD_RUN := viscosityTON.Q AND PASTE_E_STOP_NC;

IF VFD_RUN THEN
    PUMP_RUNTIME_ACC := PUMP_RUNTIME_ACC + TIME_TO_LTIME(CycleTime);
END_IF;

IF PUMP_RUNTIME_ACC >= LTIME#500h THEN
    PUMP_MAINT_DUE := TRUE;
END_IF;

END_FUNCTION_BLOCK

(* ---- public-hard-03.candidate_01.st ---- *)
(* ENGINEERING_CONTRACT
   Activations: each add/delete/modify/query acted on a rising edge via R_TRIG; no edge -> all operation outputs/error/status cleared (PUB002).
   recipeAdded/recipeDeleted/recipeModified pulse TRUE on one successful edge scan only.
   error/status pulse on same scan as the request edge; status 0 on success or idle; no latch.
   recipeQueryResult zeroed except for successful query (PUB009).
   Simultaneous rising command edges: error=TRUE, status=16#8006, no database change (unspecified).
   Add: duplicate non-zero ID -> 16#8002; no empty slot -> 16#8003; else store at lowest empty index 1..10 (PUB010).
   Delete: not found -> 16#8004; else clear whole slot and set recipeID=0 (PUB011).
   Modify: not found -> 16#8005; else replace whole slot with recipeIn (PUB012).
   Query: not found -> 16#8001; else copy matched non-zero slot to result (PUB009).
   Input recipeID=0 is treated as invalid/absent: add -> 16#8002, delete/modify/query -> not found; empty slots are not considered existing recipes.
*)
(* CONTRACT_RULES [] *)

TYPE ST_Recipe :
STRUCT
    recipeID : INT;
    ingredientType : INT;
    ingredientRatio : REAL;
    productionTemperature : REAL;
END_STRUCT
END_TYPE;

FUNCTION_BLOCK FB_RecipeManagement
VAR_INPUT
    addRecipe : BOOL;
    deleteRecipe : BOOL;
    modifyRecipe : BOOL;
    queryRecipe : BOOL;
    recipeIn : ST_Recipe;
END_VAR
VAR_OUTPUT
    recipeAdded : BOOL;
    recipeDeleted : BOOL;
    recipeModified : BOOL;
    recipeQueryResult : ST_Recipe;
    error : BOOL;
    status : WORD;
END_VAR
VAR_IN_OUT
    recipe : ARRAY[1..10] OF ST_Recipe;
END_VAR
VAR
    rtrigAdd : R_TRIG;
    rtrigDelete : R_TRIG;
    rtrigModify : R_TRIG;
    rtrigQuery : R_TRIG;

    local_AddEdge : BOOL;
    local_DeleteEdge : BOOL;
    local_ModifyEdge : BOOL;
    local_QueryEdge : BOOL;
    local_commandCount : INT;
    local_idx : INT;
    local_foundIndex : INT;
    local_emptyIndex : INT;
    local_duplicateFound : BOOL;
END_VAR

rtrigAdd(CLK := addRecipe);
rtrigDelete(CLK := deleteRecipe);
rtrigModify(CLK := modifyRecipe);
rtrigQuery(CLK := queryRecipe);

local_AddEdge := rtrigAdd.Q;
local_DeleteEdge := rtrigDelete.Q;
local_ModifyEdge := rtrigModify.Q;
local_QueryEdge := rtrigQuery.Q;

recipeAdded := FALSE;
recipeDeleted := FALSE;
recipeModified := FALSE;
error := FALSE;
status := 0;
recipeQueryResult.recipeID := 0;
recipeQueryResult.ingredientType := 0;
recipeQueryResult.ingredientRatio := 0.0;
recipeQueryResult.productionTemperature := 0.0;

local_commandCount := BOOL_TO_INT(local_AddEdge) + BOOL_TO_INT(local_DeleteEdge)
                      + BOOL_TO_INT(local_ModifyEdge) + BOOL_TO_INT(local_QueryEdge);

IF local_commandCount > 1 THEN
    error := TRUE;
    status := 16#8006;
    RETURN;
END_IF;

IF local_AddEdge THEN
    IF recipeIn.recipeID = 0 THEN
        error := TRUE;
        status := 16#8002;
        RETURN;
    END_IF;

    local_duplicateFound := FALSE;
    FOR local_idx := 1 TO 10 BY 1 DO
        IF (recipe[local_idx].recipeID <> 0) AND (recipe[local_idx].recipeID = recipeIn.recipeID) THEN
            local_duplicateFound := TRUE;
            EXIT;
        END_IF;
    END_FOR;

    IF local_duplicateFound THEN
        error := TRUE;
        status := 16#8002;
    ELSE
        local_emptyIndex := 0;
        FOR local_idx := 1 TO 10 BY 1 DO
            IF recipe[local_idx].recipeID = 0 THEN
                local_emptyIndex := local_idx;
                EXIT;
            END_IF;
        END_FOR;

        IF local_emptyIndex = 0 THEN
            error := TRUE;
            status := 16#8003;
        ELSE
            recipe[local_emptyIndex] := recipeIn;
            recipeAdded := TRUE;
        END_IF;
    END_IF;

    RETURN;
END_IF;

IF local_DeleteEdge THEN
    local_foundIndex := 0;
    FOR local_idx := 1 TO 10 BY 1 DO
        IF (recipe[local_idx].recipeID <> 0) AND (recipe[local_idx].recipeID = recipeIn.recipeID) THEN
            local_foundIndex := local_idx;
            EXIT;
        END_IF;
    END_FOR;

    IF local_foundIndex = 0 THEN
        error := TRUE;
        status := 16#8004;
    ELSE
        recipe[local_foundIndex].recipeID := 0;
        recipe[local_foundIndex].ingredientType := 0;
        recipe[local_foundIndex].ingredientRatio := 0.0;
        recipe[local_foundIndex].productionTemperature := 0.0;
        recipeDeleted := TRUE;
    END_IF;

    RETURN;
END_IF;

IF local_ModifyEdge THEN
    local_foundIndex := 0;
    FOR local_idx := 1 TO 10 BY 1 DO
        IF (recipe[local_idx].recipeID <> 0) AND (recipe[local_idx].recipeID = recipeIn.recipeID) THEN
            local_foundIndex := local_idx;
            EXIT;
        END_IF;
    END_FOR;

    IF local_foundIndex = 0 THEN
        error := TRUE;
        status := 16#8005;
    ELSE
        recipe[local_foundIndex] := recipeIn;
        recipeModified := TRUE;
    END_IF;

    RETURN;
END_IF;

IF local_QueryEdge THEN
    local_foundIndex := 0;
    FOR local_idx := 1 TO 10 BY 1 DO
        IF (recipe[local_idx].recipeID <> 0) AND (recipe[local_idx].recipeID = recipeIn.recipeID) THEN
            local_foundIndex := local_idx;
            EXIT;
        END_IF;
    END_FOR;

    IF local_foundIndex = 0 THEN
        error := TRUE;
        status := 16#8001;
    ELSE
        recipeQueryResult := recipe[local_foundIndex];
    END_IF;

    RETURN;
END_IF;

END_FUNCTION_BLOCK

(* ---- public-hard-03.candidate_02.st ---- *)
(* ENGINEERING_CONTRACT
   Activations: each add/delete/modify/query acted on a rising edge via R_TRIG; no edge -> all operation outputs/error/status cleared (PUB002).
   recipeAdded/recipeDeleted/recipeModified pulse TRUE on one successful edge scan only.
   error/status pulse on same scan as the request edge; status 0 on success or idle; no latch.
   recipeQueryResult zeroed except for successful query (PUB009).
   Simultaneous rising command edges: only the highest-priority command (add > delete > modify > query) is executed; others ignored (unspecified, deterministic).
   Add: duplicate non-zero ID -> 16#8002; no empty slot -> 16#8003; else store at lowest empty index 1..10 (PUB010).
   Delete: not found -> 16#8004; else clear whole slot and set recipeID=0 (PUB011).
   Modify: not found -> 16#8005; else replace whole slot with recipeIn (PUB012).
   Query: not found -> 16#8001; else copy matched non-zero slot to result (PUB009).
   Input recipeID=0 is treated as invalid/absent: add -> 16#8002, delete/modify/query -> not found; empty slots are not considered existing recipes.
*)
(* CONTRACT_RULES [] *)

TYPE ST_Recipe :
STRUCT
    recipeID : INT;
    ingredientType : INT;
    ingredientRatio : REAL;
    productionTemperature : REAL;
END_STRUCT
END_TYPE;

FUNCTION_BLOCK FB_RecipeManagement
VAR_INPUT
    addRecipe : BOOL;
    deleteRecipe : BOOL;
    modifyRecipe : BOOL;
    queryRecipe : BOOL;
    recipeIn : ST_Recipe;
END_VAR
VAR_OUTPUT
    recipeAdded : BOOL;
    recipeDeleted : BOOL;
    recipeModified : BOOL;
    recipeQueryResult : ST_Recipe;
    error : BOOL;
    status : WORD;
END_VAR
VAR_IN_OUT
    recipe : ARRAY[1..10] OF ST_Recipe;
END_VAR
VAR
    rtrigAdd : R_TRIG;
    rtrigDelete : R_TRIG;
    rtrigModify : R_TRIG;
    rtrigQuery : R_TRIG;

    local_AddEdge : BOOL;
    local_DeleteEdge : BOOL;
    local_ModifyEdge : BOOL;
    local_QueryEdge : BOOL;
    local_idx : INT;
    local_foundIndex : INT;
    local_emptyIndex : INT;
    local_duplicateFound : BOOL;
END_VAR

rtrigAdd(CLK := addRecipe);
rtrigDelete(CLK := deleteRecipe);
rtrigModify(CLK := modifyRecipe);
rtrigQuery(CLK := queryRecipe);

local_AddEdge := rtrigAdd.Q;
local_DeleteEdge := rtrigDelete.Q;
local_ModifyEdge := rtrigModify.Q;
local_QueryEdge := rtrigQuery.Q;

recipeAdded := FALSE;
recipeDeleted := FALSE;
recipeModified := FALSE;
error := FALSE;
status := 0;
recipeQueryResult.recipeID := 0;
recipeQueryResult.ingredientType := 0;
recipeQueryResult.ingredientRatio := 0.0;
recipeQueryResult.productionTemperature := 0.0;

IF local_AddEdge THEN
    IF recipeIn.recipeID = 0 THEN
        error := TRUE;
        status := 16#8002;
    ELSE
        local_duplicateFound := FALSE;
        FOR local_idx := 1 TO 10 BY 1 DO
            IF (recipe[local_idx].recipeID <> 0) AND (recipe[local_idx].recipeID = recipeIn.recipeID) THEN
                local_duplicateFound := TRUE;
                EXIT;
            END_IF;
        END_FOR;

        IF local_duplicateFound THEN
            error := TRUE;
            status := 16#8002;
        ELSE
            local_emptyIndex := 0;
            FOR local_idx := 1 TO 10 BY 1 DO
                IF recipe[local_idx].recipeID = 0 THEN
                    local_emptyIndex := local_idx;
                    EXIT;
                END_IF;
            END_FOR;

            IF local_emptyIndex = 0 THEN
                error := TRUE;
                status := 16#8003;
            ELSE
                recipe[local_emptyIndex] := recipeIn;
                recipeAdded := TRUE;
            END_IF;
        END_IF;
    END_IF;

ELSIF local_DeleteEdge THEN
    local_foundIndex := 0;
    FOR local_idx := 1 TO 10 BY 1 DO
        IF (recipe[local_idx].recipeID <> 0) AND (recipe[local_idx].recipeID = recipeIn.recipeID) THEN
            local_foundIndex := local_idx;
            EXIT;
        END_IF;
    END_FOR;

    IF local_foundIndex = 0 THEN
        error := TRUE;
        status := 16#8004;
    ELSE
        recipe[local_foundIndex].recipeID := 0;
        recipe[local_foundIndex].ingredientType := 0;
        recipe[local_foundIndex].ingredientRatio := 0.0;
        recipe[local_foundIndex].productionTemperature := 0.0;
        recipeDeleted := TRUE;
    END_IF;

ELSIF local_ModifyEdge THEN
    local_foundIndex := 0;
    FOR local_idx := 1 TO 10 BY 1 DO
        IF (recipe[local_idx].recipeID <> 0) AND (recipe[local_idx].recipeID = recipeIn.recipeID) THEN
            local_foundIndex := local_idx;
            EXIT;
        END_IF;
    END_FOR;

    IF local_foundIndex = 0 THEN
        error := TRUE;
        status := 16#8005;
    ELSE
        recipe[local_foundIndex] := recipeIn;
        recipeModified := TRUE;
    END_IF;

ELSIF local_QueryEdge THEN
    local_foundIndex := 0;
    FOR local_idx := 1 TO 10 BY 1 DO
        IF (recipe[local_idx].recipeID <> 0) AND (recipe[local_idx].recipeID = recipeIn.recipeID) THEN
            local_foundIndex := local_idx;
            EXIT;
        END_IF;
    END_FOR;

    IF local_foundIndex = 0 THEN
        error := TRUE;
        status := 16#8001;
    ELSE
        recipeQueryResult := recipe[local_foundIndex];
    END_IF;
END_IF;

END_FUNCTION_BLOCK

(* ---- public-hard-03.candidate_03.st ---- *)
(* ENGINEERING_CONTRACT
   Activations: each add/delete/modify/query acted on a rising edge via R_TRIG; no edge -> all operation outputs/error/status cleared (PUB002).
   recipeAdded/recipeDeleted/recipeModified pulse TRUE on one successful edge scan only.
   error/status pulse on same scan as the request edge; status 0 on success or idle; no latch.
   recipeQueryResult zeroed except for successful query (PUB009).
   Simultaneous rising command edges: each command is processed sequentially in order add, delete, modify, query.
   Add: duplicate non-zero ID -> 16#8002; no empty slot -> 16#8003; else store at lowest empty index 1..10 (PUB010).
   Delete: not found -> 16#8004; else clear whole slot and set recipeID=0 (PUB011).
   Modify: not found -> 16#8005; else replace whole slot with recipeIn (PUB012).
   Query: not found -> 16#8001; else copy matched non-zero slot to result (PUB009).
   Input recipeID=0 is treated as invalid/absent: add -> 16#8002, delete/modify/query -> not found; empty slots are not considered existing recipes.
*)
(* CONTRACT_RULES [] *)

TYPE ST_Recipe :
STRUCT
    recipeID : INT;
    ingredientType : INT;
    ingredientRatio : REAL;
    productionTemperature : REAL;
END_STRUCT
END_TYPE;

FUNCTION_BLOCK FB_RecipeManagement
VAR_INPUT
    addRecipe : BOOL;
    deleteRecipe : BOOL;
    modifyRecipe : BOOL;
    queryRecipe : BOOL;
    recipeIn : ST_Recipe;
END_VAR
VAR_OUTPUT
    recipeAdded : BOOL;
    recipeDeleted : BOOL;
    recipeModified : BOOL;
    recipeQueryResult : ST_Recipe;
    error : BOOL;
    status : WORD;
END_VAR
VAR_IN_OUT
    recipe : ARRAY[1..10] OF ST_Recipe;
END_VAR
VAR
    rtrigAdd : R_TRIG;
    rtrigDelete : R_TRIG;
    rtrigModify : R_TRIG;
    rtrigQuery : R_TRIG;

    local_AddEdge : BOOL;
    local_DeleteEdge : BOOL;
    local_ModifyEdge : BOOL;
    local_QueryEdge : BOOL;
    local_idx : INT;
    local_foundIndex : INT;
    local_emptyIndex : INT;
    local_duplicateFound : BOOL;
END_VAR

rtrigAdd(CLK := addRecipe);
rtrigDelete(CLK := deleteRecipe);
rtrigModify(CLK := modifyRecipe);
rtrigQuery(CLK := queryRecipe);

local_AddEdge := rtrigAdd.Q;
local_DeleteEdge := rtrigDelete.Q;
local_ModifyEdge := rtrigModify.Q;
local_QueryEdge := rtrigQuery.Q;

recipeAdded := FALSE;
recipeDeleted := FALSE;
recipeModified := FALSE;
error := FALSE;
status := 0;
recipeQueryResult.recipeID := 0;
recipeQueryResult.ingredientType := 0;
recipeQueryResult.ingredientRatio := 0.0;
recipeQueryResult.productionTemperature := 0.0;

(* Process add request on rising edge *)
IF local_AddEdge THEN
    IF recipeIn.recipeID = 0 THEN
        error := TRUE;
        status := 16#8002;
    ELSE
        local_duplicateFound := FALSE;
        FOR local_idx := 1 TO 10 BY 1 DO
            IF (recipe[local_idx].recipeID <> 0) AND (recipe[local_idx].recipeID = recipeIn.recipeID) THEN
                local_duplicateFound := TRUE;
                EXIT;
            END_IF;
        END_FOR;

        IF local_duplicateFound THEN
            error := TRUE;
            status := 16#8002;
        ELSE
            local_emptyIndex := 0;
            FOR local_idx := 1 TO 10 BY 1 DO
                IF recipe[local_idx].recipeID = 0 THEN
                    local_emptyIndex := local_idx;
                    EXIT;
                END_IF;
            END_FOR;

            IF local_emptyIndex = 0 THEN
                error := TRUE;
                status := 16#8003;
            ELSE
                recipe[local_emptyIndex] := recipeIn;
                recipeAdded := TRUE;
            END_IF;
        END_IF;
    END_IF;
END_IF;

(* Process delete request on rising edge *)
IF local_DeleteEdge THEN
    local_foundIndex := 0;
    FOR local_idx := 1 TO 10 BY 1 DO
        IF (recipe[local_idx].recipeID <> 0) AND (recipe[local_idx].recipeID = recipeIn.recipeID) THEN
            local_foundIndex := local_idx;
            EXIT;
        END_IF;
    END_FOR;

    IF local_foundIndex = 0 THEN
        error := TRUE;
        status := 16#8004;
    ELSE
        recipe[local_foundIndex].recipeID := 0;
        recipe[local_foundIndex].ingredientType := 0;
        recipe[local_foundIndex].ingredientRatio := 0.0;
        recipe[local_foundIndex].productionTemperature := 0.0;
        recipeDeleted := TRUE;
    END_IF;
END_IF;

(* Process modify request on rising edge *)
IF local_ModifyEdge THEN
    local_foundIndex := 0;
    FOR local_idx := 1 TO 10 BY 1 DO
        IF (recipe[local_idx].recipeID <> 0) AND (recipe[local_idx].recipeID = recipeIn.recipeID) THEN
            local_foundIndex := local_idx;
            EXIT;
        END_IF;
    END_FOR;

    IF local_foundIndex = 0 THEN
        error := TRUE;
        status := 16#8005;
    ELSE
        recipe[local_foundIndex] := recipeIn;
        recipeModified := TRUE;
    END_IF;
END_IF;

(* Process query request on rising edge *)
IF local_QueryEdge THEN
    local_foundIndex := 0;
    FOR local_idx := 1 TO 10 BY 1 DO
        IF (recipe[local_idx].recipeID <> 0) AND (recipe[local_idx].recipeID = recipeIn.recipeID) THEN
            local_foundIndex := local_idx;
            EXIT;
        END_IF;
    END_FOR;

    IF local_foundIndex = 0 THEN
        error := TRUE;
        status := 16#8001;
    ELSE
        recipeQueryResult := recipe[local_foundIndex];
    END_IF;
END_IF;

END_FUNCTION_BLOCK

(* ---- public-hard-03.raw_candidate_01.st ---- *)
(* ENGINEERING_CONTRACT
   Activations: each add/delete/modify/query acted on a rising edge via R_TRIG; no edge -> all operation outputs/error/status cleared (PUB002).
   recipeAdded/recipeDeleted/recipeModified pulse TRUE on one successful edge scan only.
   error/status pulse on same scan as the request edge; status 0 on success or idle; no latch.
   recipeQueryResult zeroed except for successful query (PUB009).
   Simultaneous rising command edges: error=TRUE, status=16#8006, no database change (unspecified).
   Add: duplicate non-zero ID -> 16#8002; no empty slot -> 16#8003; else store at lowest empty index 1..10 (PUB010).
   Delete: not found -> 16#8004; else clear whole slot and set recipeID=0 (PUB011).
   Modify: not found -> 16#8005; else replace whole slot with recipeIn (PUB012).
   Query: not found -> 16#8001; else copy matched non-zero slot to result (PUB009).
   Input recipeID=0 is treated as invalid/absent: add -> 16#8002, delete/modify/query -> not found; empty slots are not considered existing recipes.
*)
(* CONTRACT_RULES [] *)

TYPE ST_Recipe :
STRUCT
    recipeID : INT;
    ingredientType : INT;
    ingredientRatio : REAL;
    productionTemperature : REAL;
END_STRUCT
END_TYPE

FUNCTION_BLOCK FB_RecipeManagement
VAR_INPUT
    addRecipe : BOOL;
    deleteRecipe : BOOL;
    modifyRecipe : BOOL;
    queryRecipe : BOOL;
    recipeIn : ST_Recipe;
END_VAR
VAR_OUTPUT
    recipeAdded : BOOL;
    recipeDeleted : BOOL;
    recipeModified : BOOL;
    recipeQueryResult : ST_Recipe;
    error : BOOL;
    status : WORD;
END_VAR
VAR_IN_OUT
    recipe : ARRAY[1..10] OF ST_Recipe;
END_VAR
VAR
    rtrigAdd : R_TRIG;
    rtrigDelete : R_TRIG;
    rtrigModify : R_TRIG;
    rtrigQuery : R_TRIG;

    local_AddEdge : BOOL;
    local_DeleteEdge : BOOL;
    local_ModifyEdge : BOOL;
    local_QueryEdge : BOOL;
    local_commandCount : INT;
    local_idx : INT;
    local_foundIndex : INT;
    local_emptyIndex : INT;
    local_duplicateFound : BOOL;
END_VAR

rtrigAdd(CLK := addRecipe);
rtrigDelete(CLK := deleteRecipe);
rtrigModify(CLK := modifyRecipe);
rtrigQuery(CLK := queryRecipe);

local_AddEdge := rtrigAdd.Q;
local_DeleteEdge := rtrigDelete.Q;
local_ModifyEdge := rtrigModify.Q;
local_QueryEdge := rtrigQuery.Q;

recipeAdded := FALSE;
recipeDeleted := FALSE;
recipeModified := FALSE;
error := FALSE;
status := 0;
recipeQueryResult.recipeID := 0;
recipeQueryResult.ingredientType := 0;
recipeQueryResult.ingredientRatio := 0.0;
recipeQueryResult.productionTemperature := 0.0;

local_commandCount := BOOL_TO_INT(local_AddEdge) + BOOL_TO_INT(local_DeleteEdge)
                      + BOOL_TO_INT(local_ModifyEdge) + BOOL_TO_INT(local_QueryEdge);

IF local_commandCount > 1 THEN
    error := TRUE;
    status := 16#8006;
    RETURN;
END_IF;

IF local_AddEdge THEN
    IF recipeIn.recipeID = 0 THEN
        error := TRUE;
        status := 16#8002;
        RETURN;
    END_IF;

    local_duplicateFound := FALSE;
    FOR local_idx := 1 TO 10 BY 1 DO
        IF (recipe[local_idx].recipeID <> 0) AND (recipe[local_idx].recipeID = recipeIn.recipeID) THEN
            local_duplicateFound := TRUE;
            EXIT;
        END_IF;
    END_FOR;

    IF local_duplicateFound THEN
        error := TRUE;
        status := 16#8002;
    ELSE
        local_emptyIndex := 0;
        FOR local_idx := 1 TO 10 BY 1 DO
            IF recipe[local_idx].recipeID = 0 THEN
                local_emptyIndex := local_idx;
                EXIT;
            END_IF;
        END_FOR;

        IF local_emptyIndex = 0 THEN
            error := TRUE;
            status := 16#8003;
        ELSE
            recipe[local_emptyIndex] := recipeIn;
            recipeAdded := TRUE;
        END_IF;
    END_IF;

    RETURN;
END_IF;

IF local_DeleteEdge THEN
    local_foundIndex := 0;
    FOR local_idx := 1 TO 10 BY 1 DO
        IF (recipe[local_idx].recipeID <> 0) AND (recipe[local_idx].recipeID = recipeIn.recipeID) THEN
            local_foundIndex := local_idx;
            EXIT;
        END_IF;
    END_FOR;

    IF local_foundIndex = 0 THEN
        error := TRUE;
        status := 16#8004;
    ELSE
        recipe[local_foundIndex].recipeID := 0;
        recipe[local_foundIndex].ingredientType := 0;
        recipe[local_foundIndex].ingredientRatio := 0.0;
        recipe[local_foundIndex].productionTemperature := 0.0;
        recipeDeleted := TRUE;
    END_IF;

    RETURN;
END_IF;

IF local_ModifyEdge THEN
    local_foundIndex := 0;
    FOR local_idx := 1 TO 10 BY 1 DO
        IF (recipe[local_idx].recipeID <> 0) AND (recipe[local_idx].recipeID = recipeIn.recipeID) THEN
            local_foundIndex := local_idx;
            EXIT;
        END_IF;
    END_FOR;

    IF local_foundIndex = 0 THEN
        error := TRUE;
        status := 16#8005;
    ELSE
        recipe[local_foundIndex] := recipeIn;
        recipeModified := TRUE;
    END_IF;

    RETURN;
END_IF;

IF local_QueryEdge THEN
    local_foundIndex := 0;
    FOR local_idx := 1 TO 10 BY 1 DO
        IF (recipe[local_idx].recipeID <> 0) AND (recipe[local_idx].recipeID = recipeIn.recipeID) THEN
            local_foundIndex := local_idx;
            EXIT;
        END_IF;
    END_FOR;

    IF local_foundIndex = 0 THEN
        error := TRUE;
        status := 16#8001;
    ELSE
        recipeQueryResult := recipe[local_foundIndex];
    END_IF;

    RETURN;
END_IF;

END_FUNCTION_BLOCK

(* ---- public-hard-03.raw_candidate_02.st ---- *)
(* ENGINEERING_CONTRACT
   Activations: each add/delete/modify/query acted on a rising edge via R_TRIG; no edge -> all operation outputs/error/status cleared (PUB002).
   recipeAdded/recipeDeleted/recipeModified pulse TRUE on one successful edge scan only.
   error/status pulse on same scan as the request edge; status 0 on success or idle; no latch.
   recipeQueryResult zeroed except for successful query (PUB009).
   Simultaneous rising command edges: only the highest-priority command (add > delete > modify > query) is executed; others ignored (unspecified, deterministic).
   Add: duplicate non-zero ID -> 16#8002; no empty slot -> 16#8003; else store at lowest empty index 1..10 (PUB010).
   Delete: not found -> 16#8004; else clear whole slot and set recipeID=0 (PUB011).
   Modify: not found -> 16#8005; else replace whole slot with recipeIn (PUB012).
   Query: not found -> 16#8001; else copy matched non-zero slot to result (PUB009).
   Input recipeID=0 is treated as invalid/absent: add -> 16#8002, delete/modify/query -> not found; empty slots are not considered existing recipes.
*)
(* CONTRACT_RULES [] *)

TYPE ST_Recipe :
STRUCT
    recipeID : INT;
    ingredientType : INT;
    ingredientRatio : REAL;
    productionTemperature : REAL;
END_STRUCT
END_TYPE;

FUNCTION_BLOCK FB_RecipeManagement
VAR_INPUT
    addRecipe : BOOL;
    deleteRecipe : BOOL;
    modifyRecipe : BOOL;
    queryRecipe : BOOL;
    recipeIn : ST_Recipe;
END_VAR
VAR_OUTPUT
    recipeAdded : BOOL;
    recipeDeleted : BOOL;
    recipeModified : BOOL;
    recipeQueryResult : ST_Recipe;
    error : BOOL;
    status : WORD;
END_VAR
VAR_IN_OUT
    recipe : ARRAY[1..10] OF ST_Recipe;
END_VAR
VAR
    rtrigAdd : R_TRIG;
    rtrigDelete : R_TRIG;
    rtrigModify : R_TRIG;
    rtrigQuery : R_TRIG;

    local_AddEdge : BOOL;
    local_DeleteEdge : BOOL;
    local_ModifyEdge : BOOL;
    local_QueryEdge : BOOL;
    local_idx : INT;
    local_foundIndex : INT;
    local_emptyIndex : INT;
    local_duplicateFound : BOOL;
END_VAR

rtrigAdd(CLK := addRecipe);
rtrigDelete(CLK := deleteRecipe);
rtrigModify(CLK := modifyRecipe);
rtrigQuery(CLK := queryRecipe);

local_AddEdge := rtrigAdd.Q;
local_DeleteEdge := rtrigDelete.Q;
local_ModifyEdge := rtrigModify.Q;
local_QueryEdge := rtrigQuery.Q;

recipeAdded := FALSE;
recipeDeleted := FALSE;
recipeModified := FALSE;
error := FALSE;
status := 0;
recipeQueryResult.recipeID := 0;
recipeQueryResult.ingredientType := 0;
recipeQueryResult.ingredientRatio := 0.0;
recipeQueryResult.productionTemperature := 0.0;

IF local_AddEdge THEN
    IF recipeIn.recipeID = 0 THEN
        error := TRUE;
        status := 16#8002;
    ELSE
        local_duplicateFound := FALSE;
        FOR local_idx := 1 TO 10 BY 1 DO
            IF (recipe[local_idx].recipeID <> 0) AND (recipe[local_idx].recipeID = recipeIn.recipeID) THEN
                local_duplicateFound := TRUE;
                EXIT;
            END_IF;
        END_FOR;

        IF local_duplicateFound THEN
            error := TRUE;
            status := 16#8002;
        ELSE
            local_emptyIndex := 0;
            FOR local_idx := 1 TO 10 BY 1 DO
                IF recipe[local_idx].recipeID = 0 THEN
                    local_emptyIndex := local_idx;
                    EXIT;
                END_IF;
            END_FOR;

            IF local_emptyIndex = 0 THEN
                error := TRUE;
                status := 16#8003;
            ELSE
                recipe[local_emptyIndex] := recipeIn;
                recipeAdded := TRUE;
            END_IF;
        END_IF;
    END_IF;

ELSIF local_DeleteEdge THEN
    local_foundIndex := 0;
    FOR local_idx := 1 TO 10 BY 1 DO
        IF (recipe[local_idx].recipeID <> 0) AND (recipe[local_idx].recipeID = recipeIn.recipeID) THEN
            local_foundIndex := local_idx;
            EXIT;
        END_IF;
    END_FOR;

    IF local_foundIndex = 0 THEN
        error := TRUE;
        status := 16#8004;
    ELSE
        recipe[local_foundIndex].recipeID := 0;
        recipe[local_foundIndex].ingredientType := 0;
        recipe[local_foundIndex].ingredientRatio := 0.0;
        recipe[local_foundIndex].productionTemperature := 0.0;
        recipeDeleted := TRUE;
    END_IF;

ELSIF local_ModifyEdge THEN
    local_foundIndex := 0;
    FOR local_idx := 1 TO 10 BY 1 DO
        IF (recipe[local_idx].recipeID <> 0) AND (recipe[local_idx].recipeID = recipeIn.recipeID) THEN
            local_foundIndex := local_idx;
            EXIT;
        END_IF;
    END_FOR;

    IF local_foundIndex = 0 THEN
        error := TRUE;
        status := 16#8005;
    ELSE
        recipe[local_foundIndex] := recipeIn;
        recipeModified := TRUE;
    END_IF;

ELSIF local_QueryEdge THEN
    local_foundIndex := 0;
    FOR local_idx := 1 TO 10 BY 1 DO
        IF (recipe[local_idx].recipeID <> 0) AND (recipe[local_idx].recipeID = recipeIn.recipeID) THEN
            local_foundIndex := local_idx;
            EXIT;
        END_IF;
    END_FOR;

    IF local_foundIndex = 0 THEN
        error := TRUE;
        status := 16#8001;
    ELSE
        recipeQueryResult := recipe[local_foundIndex];
    END_IF;
END_IF;

END_FUNCTION_BLOCK

(* ---- public-hard-03.raw_candidate_03.st ---- *)
(* ENGINEERING_CONTRACT
   Activations: each add/delete/modify/query acted on a rising edge via R_TRIG; no edge -> all operation outputs/error/status cleared (PUB002).
   recipeAdded/recipeDeleted/recipeModified pulse TRUE on one successful edge scan only.
   error/status pulse on same scan as the request edge; status 0 on success or idle; no latch.
   recipeQueryResult zeroed except for successful query (PUB009).
   Simultaneous rising command edges: each command is processed sequentially in order add, delete, modify, query.
   Add: duplicate non-zero ID -> 16#8002; no empty slot -> 16#8003; else store at lowest empty index 1..10 (PUB010).
   Delete: not found -> 16#8004; else clear whole slot and set recipeID=0 (PUB011).
   Modify: not found -> 16#8005; else replace whole slot with recipeIn (PUB012).
   Query: not found -> 16#8001; else copy matched non-zero slot to result (PUB009).
   Input recipeID=0 is treated as invalid/absent: add -> 16#8002, delete/modify/query -> not found; empty slots are not considered existing recipes.
*)
(* CONTRACT_RULES [] *)

TYPE ST_Recipe :
STRUCT
    recipeID : INT;
    ingredientType : INT;
    ingredientRatio : REAL;
    productionTemperature : REAL;
END_STRUCT
END_TYPE;

FUNCTION_BLOCK FB_RecipeManagement
VAR_INPUT
    addRecipe : BOOL;
    deleteRecipe : BOOL;
    modifyRecipe : BOOL;
    queryRecipe : BOOL;
    recipeIn : ST_Recipe;
END_VAR
VAR_OUTPUT
    recipeAdded : BOOL;
    recipeDeleted : BOOL;
    recipeModified : BOOL;
    recipeQueryResult : ST_Recipe;
    error : BOOL;
    status : WORD;
END_VAR
VAR_IN_OUT
    recipe : ARRAY[1..10] OF ST_Recipe;
END_VAR
VAR
    rtrigAdd : R_TRIG;
    rtrigDelete : R_TRIG;
    rtrigModify : R_TRIG;
    rtrigQuery : R_TRIG;

    local_AddEdge : BOOL;
    local_DeleteEdge : BOOL;
    local_ModifyEdge : BOOL;
    local_QueryEdge : BOOL;
    local_idx : INT;
    local_foundIndex : INT;
    local_emptyIndex : INT;
    local_duplicateFound : BOOL;
END_VAR

rtrigAdd(CLK := addRecipe);
rtrigDelete(CLK := deleteRecipe);
rtrigModify(CLK := modifyRecipe);
rtrigQuery(CLK := queryRecipe);

local_AddEdge := rtrigAdd.Q;
local_DeleteEdge := rtrigDelete.Q;
local_ModifyEdge := rtrigModify.Q;
local_QueryEdge := rtrigQuery.Q;

recipeAdded := FALSE;
recipeDeleted := FALSE;
recipeModified := FALSE;
error := FALSE;
status := 0;
recipeQueryResult.recipeID := 0;
recipeQueryResult.ingredientType := 0;
recipeQueryResult.ingredientRatio := 0.0;
recipeQueryResult.productionTemperature := 0.0;

(* Process add request on rising edge *)
IF local_AddEdge THEN
    IF recipeIn.recipeID = 0 THEN
        error := TRUE;
        status := 16#8002;
    ELSE
        local_duplicateFound := FALSE;
        FOR local_idx := 1 TO 10 BY 1 DO
            IF (recipe[local_idx].recipeID <> 0) AND (recipe[local_idx].recipeID = recipeIn.recipeID) THEN
                local_duplicateFound := TRUE;
                EXIT;
            END_IF;
        END_FOR;

        IF local_duplicateFound THEN
            error := TRUE;
            status := 16#8002;
        ELSE
            local_emptyIndex := 0;
            FOR local_idx := 1 TO 10 BY 1 DO
                IF recipe[local_idx].recipeID = 0 THEN
                    local_emptyIndex := local_idx;
                    EXIT;
                END_IF;
            END_FOR;

            IF local_emptyIndex = 0 THEN
                error := TRUE;
                status := 16#8003;
            ELSE
                recipe[local_emptyIndex] := recipeIn;
                recipeAdded := TRUE;
            END_IF;
        END_IF;
    END_IF;
END_IF;

(* Process delete request on rising edge *)
IF local_DeleteEdge THEN
    local_foundIndex := 0;
    FOR local_idx := 1 TO 10 BY 1 DO
        IF (recipe[local_idx].recipeID <> 0) AND (recipe[local_idx].recipeID = recipeIn.recipeID) THEN
            local_foundIndex := local_idx;
            EXIT;
        END_IF;
    END_FOR;

    IF local_foundIndex = 0 THEN
        error := TRUE;
        status := 16#8004;
    ELSE
        recipe[local_foundIndex].recipeID := 0;
        recipe[local_foundIndex].ingredientType := 0;
        recipe[local_foundIndex].ingredientRatio := 0.0;
        recipe[local_foundIndex].productionTemperature := 0.0;
        recipeDeleted := TRUE;
    END_IF;
END_IF;

(* Process modify request on rising edge *)
IF local_ModifyEdge THEN
    local_foundIndex := 0;
    FOR local_idx := 1 TO 10 BY 1 DO
        IF (recipe[local_idx].recipeID <> 0) AND (recipe[local_idx].recipeID = recipeIn.recipeID) THEN
            local_foundIndex := local_idx;
            EXIT;
        END_IF;
    END_FOR;

    IF local_foundIndex = 0 THEN
        error := TRUE;
        status := 16#8005;
    ELSE
        recipe[local_foundIndex] := recipeIn;
        recipeModified := TRUE;
    END_IF;
END_IF;

(* Process query request on rising edge *)
IF local_QueryEdge THEN
    local_foundIndex := 0;
    FOR local_idx := 1 TO 10 BY 1 DO
        IF (recipe[local_idx].recipeID <> 0) AND (recipe[local_idx].recipeID = recipeIn.recipeID) THEN
            local_foundIndex := local_idx;
            EXIT;
        END_IF;
    END_FOR;

    IF local_foundIndex = 0 THEN
        error := TRUE;
        status := 16#8001;
    ELSE
        recipeQueryResult := recipe[local_foundIndex];
    END_IF;
END_IF;

END_FUNCTION_BLOCK

(* ---- public-medium-03.candidate_01.st ---- *)
FUNCTION_BLOCK FB
VAR_INPUT
    cyclicExecution : BOOL;
    trigger : BOOL;
    value : LREAL;
    windowSize : INT;
    reset : BOOL;
END_VAR
VAR_OUTPUT
    average : LREAL;
    windowSizeReached : BOOL;
    error : BOOL;
    status : WORD;
END_VAR
VAR
    tmp_trig : R_TRIG;
    local_data : ARRAY[0..99] OF LREAL;
    local_count : INT := 0;
    local_start : INT := 0;
    local_sum_all : LREAL := 0.0;
    local_avg_sum : LREAL;
    local_effective : INT;
    tmp_i : INT;
    tmp_idx : INT;
END_VAR

(* ENGINEERING_CONTRACT
 * average: updated after each accepted sample (PUB001-PUB003); on reset := 0.0; on invalid window holds last value; 0.0 until first sample.
 * windowSizeReached: TRUE when stored sample count >= windowSize (PUB001); FALSE on reset and invalid window.
 * error/status: error=TRUE, status=WORD#16#8200 when windowSize<1 or >100 (PUB004, PUB006, PUB007); reset with valid window clears to FALSE/WORD#16#0000.
 * sample priority per scan: reset first, invalid-window block second, cyclicExecution TRUE (PUB002) third, trigger rising edge (PUB003) fourth; trigger ignored while cyclicExecution TRUE.
 * reset: clears count, ring start, sum, average, and reached state (PUB004).
 * state: ring of up to 100 LREAL samples with total sum; invalid window pauses sampling and does not clear history; dynamic window changes average over last windowSize samples (unspecified by task).
 * boundaries: valid windowSize 1..100 inclusive; average shares value units; status codes match PUB006/PUB007.
 *)

(* CONTRACT_RULES [] *)

tmp_trig(CLK := trigger);

IF reset THEN
    local_count := 0;
    local_start := 0;
    local_sum_all := 0.0;
    average := 0.0;
    windowSizeReached := FALSE;
END_IF;

IF (windowSize < 1) OR (windowSize > 100) THEN
    error := TRUE;
    status := WORD#16#8200;
    windowSizeReached := FALSE;
    RETURN;
ELSE
    error := FALSE;
    status := WORD#16#0000;
END_IF;

IF reset THEN
    RETURN;
END_IF;

IF cyclicExecution THEN
    IF local_count < 100 THEN
        local_data[local_count] := value;
        local_count := local_count + 1;
        local_sum_all := local_sum_all + value;
    ELSE
        local_sum_all := local_sum_all - local_data[local_start] + value;
        local_data[local_start] := value;
        local_start := (local_start + 1) MOD 100;
    END_IF;
ELSIF tmp_trig.Q THEN
    IF local_count < 100 THEN
        local_data[local_count] := value;
        local_count := local_count + 1;
        local_sum_all := local_sum_all + value;
    ELSE
        local_sum_all := local_sum_all - local_data[local_start] + value;
        local_data[local_start] := value;
        local_start := (local_start + 1) MOD 100;
    END_IF;
END_IF;

local_avg_sum := local_sum_all;

IF local_count > windowSize THEN
    FOR tmp_i := 0 TO (local_count - windowSize - 1) DO
        tmp_idx := (local_start + tmp_i) MOD 100;
        local_avg_sum := local_avg_sum - local_data[tmp_idx];
    END_FOR;
END_IF;

local_effective := local_count;
IF local_effective > windowSize THEN
    local_effective := windowSize;
END_IF;

IF local_effective > 0 THEN
    average := local_avg_sum / INT_TO_LREAL(local_effective);
ELSE
    average := 0.0;
END_IF;

windowSizeReached := local_count >= windowSize;

END_FUNCTION_BLOCK

(* ---- public-medium-03.candidate_02.st ---- *)
FUNCTION_BLOCK FB
VAR_INPUT
    cyclicExecution : BOOL;
    trigger : BOOL;
    value : LREAL;
    windowSize : INT;
    reset : BOOL;
END_VAR
VAR_OUTPUT
    average : LREAL;
    windowSizeReached : BOOL;
    error : BOOL;
    status : WORD;
END_VAR
VAR
    tmp_trig : R_TRIG;
    local_data : ARRAY[0..99] OF LREAL;
    local_count : INT := 0;
    local_start : INT := 0;
    local_sum_all : LREAL := 0.0;
    local_avg_sum : LREAL;
    local_effective : INT;
    tmp_i : INT;
    tmp_idx : INT;
END_VAR

(* ENGINEERING_CONTRACT
 * average: updated after each accepted sample (PUB001-PUB003); on reset := 0.0; on invalid window holds last value; 0.0 until first sample.
 * windowSizeReached: TRUE when stored sample count >= windowSize (PUB001); FALSE on reset and invalid window.
 * error/status: error=TRUE, status=WORD#16#8200 when windowSize<1 or >100 (PUB004, PUB006, PUB007); reset with valid window clears to FALSE/WORD#16#0000.
 * sample priority per scan: reset first, invalid-window block second, cyclicExecution TRUE (PUB002) third, trigger rising edge (PUB003) fourth; trigger ignored while cyclicExecution TRUE.
 * reset: clears count, ring start, sum, average, and reached state (PUB004). Same-scan reset blocks any new sample to guarantee average resets to 0.0.
 * state: ring of up to 100 LREAL samples with total sum; invalid window pauses sampling and does not clear history; dynamic window changes average over last windowSize samples (unspecified by task).
 * boundaries: valid windowSize 1..100 inclusive; average shares value units; status codes match PUB006/PUB007.
 *)

(* CONTRACT_RULES [] *)

tmp_trig(CLK := trigger);

IF reset THEN
    local_count := 0;
    local_start := 0;
    local_sum_all := 0.0;
    average := 0.0;
    windowSizeReached := FALSE;
END_IF;

IF (windowSize < 1) OR (windowSize > 100) THEN
    error := TRUE;
    status := WORD#16#8200;
    windowSizeReached := FALSE;
    RETURN;
ELSE
    error := FALSE;
    status := WORD#16#0000;
END_IF;

IF reset THEN
    RETURN;
END_IF;

IF cyclicExecution THEN
    IF local_count < 100 THEN
        local_data[local_count] := value;
        local_count := local_count + 1;
        local_sum_all := local_sum_all + value;
    ELSE
        local_sum_all := local_sum_all - local_data[local_start] + value;
        local_data[local_start] := value;
        local_start := (local_start + 1) MOD 100;
    END_IF;
ELSIF tmp_trig.Q THEN
    IF local_count < 100 THEN
        local_data[local_count] := value;
        local_count := local_count + 1;
        local_sum_all := local_sum_all + value;
    ELSE
        local_sum_all := local_sum_all - local_data[local_start] + value;
        local_data[local_start] := value;
        local_start := (local_start + 1) MOD 100;
    END_IF;
END_IF;

local_avg_sum := local_sum_all;

IF local_count > windowSize THEN
    FOR tmp_i := 0 TO (local_count - windowSize - 1) DO
        tmp_idx := (local_start + tmp_i) MOD 100;
        local_avg_sum := local_avg_sum - local_data[tmp_idx];
    END_FOR;
END_IF;

local_effective := local_count;
IF local_effective > windowSize THEN
    local_effective := windowSize;
END_IF;

IF local_effective > 0 THEN
    average := local_avg_sum / INT_TO_LREAL(local_effective);
ELSE
    average := 0.0;
END_IF;

windowSizeReached := local_count >= windowSize;

END_FUNCTION_BLOCK

(* ---- public-medium-03.candidate_03.st ---- *)
FUNCTION_BLOCK FB
VAR_INPUT
    cyclicExecution : BOOL;
    trigger : BOOL;
    value : LREAL;
    windowSize : INT;
    reset : BOOL;
END_VAR
VAR_OUTPUT
    average : LREAL;
    windowSizeReached : BOOL;
    error : BOOL;
    status : WORD;
END_VAR
VAR
    tmp_trig : R_TRIG;
    local_data : ARRAY[0..99] OF LREAL;
    local_count : INT := 0;
    local_start : INT := 0;
    local_sum_all : LREAL := 0.0;
    local_avg_sum : LREAL;
    local_effective : INT;
    tmp_i : INT;
    tmp_idx : INT;
END_VAR

(* ENGINEERING_CONTRACT
 * average: updated after each accepted sample (PUB001-PUB003); 0.0 until first sample.
 * On reset: history is cleared, average assigned 0.0 and windowSizeReached FALSE.
 * If cyclicExecution is TRUE in the same scan as reset, the current value is then accepted
 * as the first sample of the new window (PUB002). If cyclicExecution is FALSE and a trigger
 * rising edge occurs in the same scan as reset, the current value is accepted (PUB003).
 * windowSizeReached: TRUE when stored sample count >= windowSize (PUB001); cleared on reset
 * and on invalid window.
 * error/status: error=TRUE, status=WORD#16#8200 when windowSize<1 or >100 (PUB004, PUB007);
 * reset with valid window clears to FALSE/WORD#16#0000.
 * sample priority per scan: reset first, invalid-window block second, cyclicExecution TRUE
 * third, trigger rising edge fourth; trigger ignored while cyclicExecution TRUE.
 * state: ring of up to 100 LREAL samples with total sum; invalid window pauses sampling and
 * does not clear history; dynamic window changes average over last windowSize samples.
 * boundaries: valid windowSize 1..100 inclusive; average shares value units.
 *)

(* CONTRACT_RULES [] *)

tmp_trig(CLK := trigger);

IF reset THEN
    local_count := 0;
    local_start := 0;
    local_sum_all := 0.0;
    average := 0.0;
    windowSizeReached := FALSE;
END_IF;

IF (windowSize < 1) OR (windowSize > 100) THEN
    error := TRUE;
    status := WORD#16#8200;
    windowSizeReached := FALSE;
    RETURN;
ELSE
    error := FALSE;
    status := WORD#16#0000;
END_IF;

IF cyclicExecution THEN
    IF local_count < 100 THEN
        local_data[local_count] := value;
        local_count := local_count + 1;
        local_sum_all := local_sum_all + value;
    ELSE
        local_sum_all := local_sum_all - local_data[local_start] + value;
        local_data[local_start] := value;
        local_start := (local_start + 1) MOD 100;
    END_IF;
ELSIF tmp_trig.Q THEN
    IF local_count < 100 THEN
        local_data[local_count] := value;
        local_count := local_count + 1;
        local_sum_all := local_sum_all + value;
    ELSE
        local_sum_all := local_sum_all - local_data[local_start] + value;
        local_data[local_start] := value;
        local_start := (local_start + 1) MOD 100;
    END_IF;
END_IF;

local_avg_sum := local_sum_all;

IF local_count > windowSize THEN
    FOR tmp_i := 0 TO (local_count - windowSize - 1) DO
        tmp_idx := (local_start + tmp_i) MOD 100;
        local_avg_sum := local_avg_sum - local_data[tmp_idx];
    END_FOR;
END_IF;

local_effective := local_count;
IF local_effective > windowSize THEN
    local_effective := windowSize;
END_IF;

IF local_effective > 0 THEN
    average := local_avg_sum / INT_TO_LREAL(local_effective);
ELSE
    average := 0.0;
END_IF;

windowSizeReached := local_count >= windowSize;

END_FUNCTION_BLOCK

(* ---- public-medium-03.candidate_04.st ---- *)
FUNCTION_BLOCK FB
VAR_INPUT
    cyclicExecution : BOOL;
    trigger : BOOL;
    value : LREAL;
    windowSize : INT;
    reset : BOOL;
END_VAR
VAR_OUTPUT
    average : LREAL;
    windowSizeReached : BOOL;
    error : BOOL;
    status : WORD;
END_VAR
VAR
    tmp_trig : R_TRIG;
    local_data : ARRAY[0..99] OF LREAL;
    local_count : INT := 0;
    local_start : INT := 0;
    local_sum_all : LREAL := 0.0;
    local_avg_sum : LREAL;
    local_effective : INT;
    tmp_i : INT;
    tmp_idx : INT;
END_VAR

(* ENGINEERING_CONTRACT
 * average: 0.0 after reset; updated after each accepted sample (PUB001-PUB003);
 *          retains last value while windowSize is invalid (unspecified in PUB004).
 * windowSizeReached: TRUE when stored sample count >= windowSize (PUB001);
 *                    FALSE on reset and while windowSize invalid.
 * error/status: error=TRUE, status=WORD#16#8200 when windowSize<1 or >100
 *               (PUB004,PUB006,PUB007); reset with valid window clears to FALSE/WORD#16#0000.
 * priority per scan: 1) validate window, 2) reset, 3) cyclicExecution, 4) trigger rising edge;
 *                   trigger ignored while cyclicExecution TRUE (interface definition).
 * reset: clears ring count, ring start, sum, average, and reached state (PUB004).
 * ring: fixed 100-slot LREAL buffer with total sum; dynamic window uses last windowSize samples.
 * boundaries: valid windowSize 1..100 inclusive; average shares value units.
 *)

(* CONTRACT_RULES [] *)

IF (windowSize < 1) OR (windowSize > 100) THEN
    error := TRUE;
    status := WORD#16#8200;
    windowSizeReached := FALSE;
    RETURN;
ELSE
    error := FALSE;
    status := WORD#16#0000;
END_IF;

IF reset THEN
    local_count := 0;
    local_start := 0;
    local_sum_all := 0.0;
    average := 0.0;
    windowSizeReached := FALSE;
    RETURN;
END_IF;

tmp_trig(CLK := trigger);

IF cyclicExecution THEN
    IF local_count < 100 THEN
        local_data[local_count] := value;
        local_count := local_count + 1;
        local_sum_all := local_sum_all + value;
    ELSE
        local_sum_all := local_sum_all - local_data[local_start] + value;
        local_data[local_start] := value;
        local_start := (local_start + 1) MOD 100;
    END_IF;
ELSIF tmp_trig.Q THEN
    IF local_count < 100 THEN
        local_data[local_count] := value;
        local_count := local_count + 1;
        local_sum_all := local_sum_all + value;
    ELSE
        local_sum_all := local_sum_all - local_data[local_start] + value;
        local_data[local_start] := value;
        local_start := (local_start + 1) MOD 100;
    END_IF;
END_IF;

local_avg_sum := local_sum_all;

IF local_count > windowSize THEN
    FOR tmp_i := 0 TO (local_count - windowSize - 1) DO
        tmp_idx := (local_start + tmp_i) MOD 100;
        local_avg_sum := local_avg_sum - local_data[tmp_idx];
    END_FOR;
END_IF;

local_effective := local_count;
IF local_effective > windowSize THEN
    local_effective := windowSize;
END_IF;

IF local_effective > 0 THEN
    average := local_avg_sum / INT_TO_LREAL(local_effective);
ELSE
    average := 0.0;
END_IF;

windowSizeReached := local_count >= windowSize;

END_FUNCTION_BLOCK

(* ---- public-medium-03.raw_candidate_01.st ---- *)
FUNCTION_BLOCK FB
VAR_INPUT
    cyclicExecution : BOOL;
    trigger : BOOL;
    value : LREAL;
    windowSize : INT;
    reset : BOOL;
END_VAR
VAR_OUTPUT
    average : LREAL;
    windowSizeReached : BOOL;
    error : BOOL;
    status : WORD;
END_VAR
VAR
    tmp_trig : R_TRIG;
    local_data : ARRAY[0..99] OF LREAL;
    local_count : INT := 0;
    local_start : INT := 0;
    local_sum_all : LREAL := 0.0;
    local_avg_sum : LREAL;
    local_effective : INT;
    tmp_i : INT;
    tmp_idx : INT;
END_VAR

(* ENGINEERING_CONTRACT
 * average: updated after each accepted sample (PUB001-PUB003); on reset := 0.0; on invalid window holds last value; 0.0 until first sample.
 * windowSizeReached: TRUE when stored sample count >= windowSize (PUB001); FALSE on reset and invalid window.
 * error/status: error=TRUE, status=WORD#16#8200 when windowSize<1 or >100 (PUB004, PUB006, PUB007); reset with valid window clears to FALSE/WORD#16#0000.
 * sample priority per scan: reset first, invalid-window block second, cyclicExecution TRUE (PUB002) third, trigger rising edge (PUB003) fourth; trigger ignored while cyclicExecution TRUE.
 * reset: clears count, ring start, sum, average, and reached state (PUB004).
 * state: ring of up to 100 LREAL samples with total sum; invalid window pauses sampling and does not clear history; dynamic window changes average over last windowSize samples (unspecified by task).
 * boundaries: valid windowSize 1..100 inclusive; average shares value units; status codes match PUB006/PUB007.
 *)

(* CONTRACT_RULES [] *)

tmp_trig(CLK := trigger);

IF reset THEN
    local_count := 0;
    local_start := 0;
    local_sum_all := 0.0;
    average := 0.0;
    windowSizeReached := FALSE;
END_IF;

IF (windowSize < 1) OR (windowSize > 100) THEN
    error := TRUE;
    status := WORD#16#8200;
    windowSizeReached := FALSE;
    RETURN;
ELSE
    error := FALSE;
    status := WORD#16#0000;
END_IF;

IF reset THEN
    RETURN;
END_IF;

IF cyclicExecution THEN
    IF local_count < 100 THEN
        local_data[local_count] := value;
        local_count := local_count + 1;
        local_sum_all := local_sum_all + value;
    ELSE
        local_sum_all := local_sum_all - local_data[local_start] + value;
        local_data[local_start] := value;
        local_start := (local_start + 1) MOD 100;
    END_IF;
ELSIF tmp_trig.Q THEN
    IF local_count < 100 THEN
        local_data[local_count] := value;
        local_count := local_count + 1;
        local_sum_all := local_sum_all + value;
    ELSE
        local_sum_all := local_sum_all - local_data[local_start] + value;
        local_data[local_start] := value;
        local_start := (local_start + 1) MOD 100;
    END_IF;
END_IF;

local_avg_sum := local_sum_all;

IF local_count > windowSize THEN
    FOR tmp_i := 0 TO (local_count - windowSize - 1) DO
        tmp_idx := (local_start + tmp_i) MOD 100;
        local_avg_sum := local_avg_sum - local_data[tmp_idx];
    END_FOR;
END_IF;

local_effective := local_count;
IF local_effective > windowSize THEN
    local_effective := windowSize;
END_IF;

IF local_effective > 0 THEN
    average := local_avg_sum / INT_TO_LREAL(local_effective);
ELSE
    average := 0.0;
END_IF;

windowSizeReached := local_count >= windowSize;

END_FUNCTION_BLOCK

(* ---- public-medium-03.raw_candidate_02.st ---- *)
FUNCTION_BLOCK FB
VAR_INPUT
    cyclicExecution : BOOL;
    trigger : BOOL;
    value : LREAL;
    windowSize : INT;
    reset : BOOL;
END_VAR
VAR_OUTPUT
    average : LREAL;
    windowSizeReached : BOOL;
    error : BOOL;
    status : WORD;
END_VAR
VAR
    tmp_trig : R_TRIG;
    local_data : ARRAY[0..99] OF LREAL;
    local_count : INT := 0;
    local_start : INT := 0;
    local_sum_all : LREAL := 0.0;
    local_avg_sum : LREAL;
    local_effective : INT;
    tmp_i : INT;
    tmp_idx : INT;
END_VAR

(* ENGINEERING_CONTRACT
 * average: updated after each accepted sample (PUB001-PUB003); on reset := 0.0; on invalid window holds last value; 0.0 until first sample.
 * windowSizeReached: TRUE when stored sample count >= windowSize (PUB001); FALSE on reset and invalid window.
 * error/status: error=TRUE, status=WORD#16#8200 when windowSize<1 or >100 (PUB004, PUB006, PUB007); reset with valid window clears to FALSE/WORD#16#0000.
 * sample priority per scan: reset first, invalid-window block second, cyclicExecution TRUE (PUB002) third, trigger rising edge (PUB003) fourth; trigger ignored while cyclicExecution TRUE.
 * reset: clears count, ring start, sum, average, and reached state (PUB004). Same-scan reset blocks any new sample to guarantee average resets to 0.0.
 * state: ring of up to 100 LREAL samples with total sum; invalid window pauses sampling and does not clear history; dynamic window changes average over last windowSize samples (unspecified by task).
 * boundaries: valid windowSize 1..100 inclusive; average shares value units; status codes match PUB006/PUB007.
 *)

(* CONTRACT_RULES [] *)

tmp_trig(CLK := trigger);

IF reset THEN
    local_count := 0;
    local_start := 0;
    local_sum_all := 0.0;
    average := 0.0;
    windowSizeReached := FALSE;
END_IF;

IF (windowSize < 1) OR (windowSize > 100) THEN
    error := TRUE;
    status := WORD#16#8200;
    windowSizeReached := FALSE;
    RETURN;
ELSE
    error := FALSE;
    status := WORD#16#0000;
END_IF;

IF reset THEN
    RETURN;
END_IF;

IF cyclicExecution THEN
    IF local_count < 100 THEN
        local_data[local_count] := value;
        local_count := local_count + 1;
        local_sum_all := local_sum_all + value;
    ELSE
        local_sum_all := local_sum_all - local_data[local_start] + value;
        local_data[local_start] := value;
        local_start := (local_start + 1) MOD 100;
    END_IF;
ELSIF tmp_trig.Q THEN
    IF local_count < 100 THEN
        local_data[local_count] := value;
        local_count := local_count + 1;
        local_sum_all := local_sum_all + value;
    ELSE
        local_sum_all := local_sum_all - local_data[local_start] + value;
        local_data[local_start] := value;
        local_start := (local_start + 1) MOD 100;
    END_IF;
END_IF;

local_avg_sum := local_sum_all;

IF local_count > windowSize THEN
    FOR tmp_i := 0 TO (local_count - windowSize - 1) DO
        tmp_idx := (local_start + tmp_i) MOD 100;
        local_avg_sum := local_avg_sum - local_data[tmp_idx];
    END_FOR;
END_IF;

local_effective := local_count;
IF local_effective > windowSize THEN
    local_effective := windowSize;
END_IF;

IF local_effective > 0 THEN
    average := local_avg_sum / INT_TO_LREAL(local_effective);
ELSE
    average := 0.0;
END_IF;

windowSizeReached := local_count >= windowSize;

END_FUNCTION_BLOCK

(* ---- public-medium-03.raw_candidate_03.st ---- *)
FUNCTION_BLOCK FB
VAR_INPUT
    cyclicExecution : BOOL;
    trigger : BOOL;
    value : LREAL;
    windowSize : INT;
    reset : BOOL;
END_VAR
VAR_OUTPUT
    average : LREAL;
    windowSizeReached : BOOL;
    error : BOOL;
    status : WORD;
END_VAR
VAR
    tmp_trig : R_TRIG;
    local_data : ARRAY[0..99] OF LREAL;
    local_count : INT := 0;
    local_start : INT := 0;
    local_sum_all : LREAL := 0.0;
    local_avg_sum : LREAL;
    local_effective : INT;
    tmp_i : INT;
    tmp_idx : INT;
END_VAR

(* ENGINEERING_CONTRACT
 * average: updated after each accepted sample (PUB001-PUB003); 0.0 until first sample.
 * On reset: history is cleared, average assigned 0.0 and windowSizeReached FALSE.
 * If cyclicExecution is TRUE in the same scan as reset, the current value is then accepted
 * as the first sample of the new window (PUB002). If cyclicExecution is FALSE and a trigger
 * rising edge occurs in the same scan as reset, the current value is accepted (PUB003).
 * windowSizeReached: TRUE when stored sample count >= windowSize (PUB001); cleared on reset
 * and on invalid window.
 * error/status: error=TRUE, status=WORD#16#8200 when windowSize<1 or >100 (PUB004, PUB007);
 * reset with valid window clears to FALSE/WORD#16#0000.
 * sample priority per scan: reset first, invalid-window block second, cyclicExecution TRUE
 * third, trigger rising edge fourth; trigger ignored while cyclicExecution TRUE.
 * state: ring of up to 100 LREAL samples with total sum; invalid window pauses sampling and
 * does not clear history; dynamic window changes average over last windowSize samples.
 * boundaries: valid windowSize 1..100 inclusive; average shares value units.
 *)

(* CONTRACT_RULES [] *)

tmp_trig(CLK := trigger);

IF reset THEN
    local_count := 0;
    local_start := 0;
    local_sum_all := 0.0;
    average := 0.0;
    windowSizeReached := FALSE;
END_IF;

IF (windowSize < 1) OR (windowSize > 100) THEN
    error := TRUE;
    status := WORD#16#8200;
    windowSizeReached := FALSE;
    RETURN;
ELSE
    error := FALSE;
    status := WORD#16#0000;
END_IF;

IF cyclicExecution THEN
    IF local_count < 100 THEN
        local_data[local_count] := value;
        local_count := local_count + 1;
        local_sum_all := local_sum_all + value;
    ELSE
        local_sum_all := local_sum_all - local_data[local_start] + value;
        local_data[local_start] := value;
        local_start := (local_start + 1) MOD 100;
    END_IF;
ELSIF tmp_trig.Q THEN
    IF local_count < 100 THEN
        local_data[local_count] := value;
        local_count := local_count + 1;
        local_sum_all := local_sum_all + value;
    ELSE
        local_sum_all := local_sum_all - local_data[local_start] + value;
        local_data[local_start] := value;
        local_start := (local_start + 1) MOD 100;
    END_IF;
END_IF;

local_avg_sum := local_sum_all;

IF local_count > windowSize THEN
    FOR tmp_i := 0 TO (local_count - windowSize - 1) DO
        tmp_idx := (local_start + tmp_i) MOD 100;
        local_avg_sum := local_avg_sum - local_data[tmp_idx];
    END_FOR;
END_IF;

local_effective := local_count;
IF local_effective > windowSize THEN
    local_effective := windowSize;
END_IF;

IF local_effective > 0 THEN
    average := local_avg_sum / INT_TO_LREAL(local_effective);
ELSE
    average := 0.0;
END_IF;

windowSizeReached := local_count >= windowSize;

END_FUNCTION_BLOCK

(* ---- public-medium-03.raw_candidate_04.st ---- *)
FUNCTION_BLOCK FB
VAR_INPUT
    cyclicExecution : BOOL;
    trigger : BOOL;
    value : LREAL;
    windowSize : INT;
    reset : BOOL;
END_VAR
VAR_OUTPUT
    average : LREAL;
    windowSizeReached : BOOL;
    error : BOOL;
    status : WORD;
END_VAR
VAR
    tmp_trig : R_TRIG;
    local_data : ARRAY[0..99] OF LREAL;
    local_count : INT := 0;
    local_start : INT := 0;
    local_sum_all : LREAL := 0.0;
    local_avg_sum : LREAL;
    local_effective : INT;
    tmp_i : INT;
    tmp_idx : INT;
END_VAR

(* ENGINEERING_CONTRACT
 * average: 0.0 after reset; updated after each accepted sample (PUB001-PUB003);
 *          retains last value while windowSize is invalid (unspecified in PUB004).
 * windowSizeReached: TRUE when stored sample count >= windowSize (PUB001);
 *                    FALSE on reset and while windowSize invalid.
 * error/status: error=TRUE, status=WORD#16#8200 when windowSize<1 or >100
 *               (PUB004,PUB006,PUB007); reset with valid window clears to FALSE/WORD#16#0000.
 * priority per scan: 1) validate window, 2) reset, 3) cyclicExecution, 4) trigger rising edge;
 *                   trigger ignored while cyclicExecution TRUE (interface definition).
 * reset: clears ring count, ring start, sum, average, and reached state (PUB004).
 * ring: fixed 100-slot LREAL buffer with total sum; dynamic window uses last windowSize samples.
 * boundaries: valid windowSize 1..100 inclusive; average shares value units.
 *)

(* CONTRACT_RULES [] *)

IF (windowSize < 1) OR (windowSize > 100) THEN
    error := TRUE;
    status := WORD#16#8200;
    windowSizeReached := FALSE;
    RETURN;
ELSE
    error := FALSE;
    status := WORD#16#0000;
END_IF;

IF reset THEN
    local_count := 0;
    local_start := 0;
    local_sum_all := 0.0;
    average := 0.0;
    windowSizeReached := FALSE;
    RETURN;
END_IF;

tmp_trig(CLK := trigger);

IF cyclicExecution THEN
    IF local_count < 100 THEN
        local_data[local_count] := value;
        local_count := local_count + 1;
        local_sum_all := local_sum_all + value;
    ELSE
        local_sum_all := local_sum_all - local_data[local_start] + value;
        local_data[local_start] := value;
        local_start := (local_start + 1) MOD 100;
    END_IF;
ELSIF tmp_trig.Q THEN
    IF local_count < 100 THEN
        local_data[local_count] := value;
        local_count := local_count + 1;
        local_sum_all := local_sum_all + value;
    ELSE
        local_sum_all := local_sum_all - local_data[local_start] + value;
        local_data[local_start] := value;
        local_start := (local_start + 1) MOD 100;
    END_IF;
END_IF;

local_avg_sum := local_sum_all;

IF local_count > windowSize THEN
    FOR tmp_i := 0 TO (local_count - windowSize - 1) DO
        tmp_idx := (local_start + tmp_i) MOD 100;
        local_avg_sum := local_avg_sum - local_data[tmp_idx];
    END_FOR;
END_IF;

local_effective := local_count;
IF local_effective > windowSize THEN
    local_effective := windowSize;
END_IF;

IF local_effective > 0 THEN
    average := local_avg_sum / INT_TO_LREAL(local_effective);
ELSE
    average := 0.0;
END_IF;

windowSizeReached := local_count >= windowSize;

END_FUNCTION_BLOCK
